(* Logix 5000 project; controller TFF vendor 1 type 14 code 107 rev 34.11; software revision 34.03; part 12 of 36 *)

        LevelConfiguration[0].Alm_HIHITMR := 2, LevelConfiguration[0].Alm_HIHITMR_PRE := 2, LevelConfiguration[1].Alm_HI := 50.0, LevelConfiguration[1].Alm_HI_PRE := 50.0, LevelConfiguration[1].Alm_HIHI := 50.0, LevelConfiguration[1].Alm_HIHI_PRE := 50.0, LevelConfiguration[1].Alm_LOLOTMR := 2, LevelConfiguration[1].Alm_LOLOTMR_PRE := 2, LevelConfiguration[1].Alm_LOTMR := 2, LevelConfiguration[1].Alm_LOTMR_PRE := 2, LevelConfiguration[1].Alm_HITMR := 2, LevelConfiguration[1].Alm_HITMR_PRE := 2, LevelConfiguration[1].Alm_HIHITMR := 2, LevelConfiguration[1].Alm_HIHITMR_PRE := 2, LevelConfiguration[2].Alm_LOLO := 20.0, LevelConfiguration[2].Alm_LOLO_PRE := 20.0, LevelConfiguration[2].Alm_LO := 40.0, LevelConfiguration[2].Alm_LO_PRE := 40.0, LevelConfiguration[2].Alm_HI := 160.0, LevelConfiguration[2].Alm_HI_PRE := 160.0, LevelConfiguration[2].Alm_HIHI := 180.0, LevelConfiguration[2].Alm_HIHI_PRE := 180.0, LevelConfiguration[2].Alm_LOLOTMR := 2, LevelConfiguration[2].Alm_LOLOTMR_PRE := 2, LevelConfiguration[2].Alm_LOTMR := 2, LevelConfiguration[2].Alm_LOTMR_PRE := 2, LevelConfiguration[2].Alm_HITMR := 2, LevelConfiguration[2].Alm_HITMR_PRE := 2, LevelConfiguration[2].Alm_HIHITMR := 2, LevelConfiguration[2].Alm_HIHITMR_PRE := 2, LevelConfiguration[3].Alm_HI := 190.0, LevelConfiguration[3].Alm_HI_PRE := 190.0, LevelConfiguration[3].Alm_HIHI := 200.0, LevelConfiguration[3].Alm_HIHI_PRE := 200.0, Feed_Bag_Tare_Timer.PRE := 3000, Filtrate_Bag_Tare_Timer.PRE := 3000);   // Tank Management
   ThisSystem : SystemType := (Value := 2, MoldType := 124, PreviousValue := 124, EnableSystemType[0] := 1, EnableSystemType[1] := 1, EnableSystemType[2] := 1, EnableSystemType[3] := 1, NewSystem_Timer.PRE := 60000, NewSystem_Timer.ACC := 177455, NewSystem_Timer.EN := 1, NewSystem_Timer.DN := 1);
   TI001 : ALIAS FOR AnalogPoint[13];   // Feed Bag Temperature
   TI001_SIG : ALIAS FOR DigitalPoint[101];
   TI001Alarm : ALIAS FOR AlarmAnalog[13];   // Feed Bag Temperature Alarm
   TimerControl : TimerControl := (Save := 20456, Seconds := 20456, Colon := ':', ColonZero := ':0', Cycle := 818248);   // Timer Control
   Timers : Timers[22] := ([0].TotalSeconds := 30.0, [0].Seconds := 30, [0].sHours := '0', [0].sMinutes := '0', [0].sSeconds := '30', [0].HMS := '0:00:30', [0].LastHMS := '0:02:09', [1].sHours := '0', [1].sMinutes := '0', [1].sSeconds := '0', [1].HMS := '0:00:00', [2].sHours := '0', [2].sMinutes := '0', [2].sSeconds := '0', [2].HMS := '0:00:00', [3].TotalSeconds := 7.0, [3].Seconds := 7, [3].sHours := '0', [3].sMinutes := '0', [3].sSeconds := '7', [3].HMS := '0:00:07', [3].LastHMS := '0:00:00', [4].TotalSeconds := 2.0, [4].Seconds := 2, [4].sHours := '0', [4].sMinutes := '0', [4].sSeconds := '2', [4].HMS := '0:00:02', [5].sHours := '0', [5].sMinutes := '0', [5].sSeconds := '0', [5].HMS := '0:00:00', [5].LastHMS := ':00$00$07$00$00$000:00:00$00$00$00$00$00$00$00$00$00$07$00$00$00', [6].sHours := '0', [6].sMinutes := '0', [6].sSeconds := '0', [6].HMS := '0:00:00', [6].LastHMS := '0:00:02', [7].sHours := '0', [7].sMinutes := '0', [7].sSeconds := '0', [7].HMS := '0:00:00', [8].sHours := '0', [8].sMinutes := '0', [8].sSeconds := '0', [8].HMS := '0:00:00', [8].LastHMS := '$07$00$00$000:00:00$00$00$00$00$00$00$00$00$00$07$00$00$000:$00$00', [9].sHours := '0', [9].sMinutes := '0', [9].sSeconds := '0', [9].HMS := '0:00:00', [9].LastHMS := '$00$00$00$00$00$00$00$00$07$00$00$000:00:00$00$07$00$00$000:$00$00', [10].sHours := '0', [10].sMinutes := '0', [10].sSeconds := '0', [10].HMS := '0:00:00', [10].LastHMS := '0:00:00', [11].sHours := '0', [11].sMinutes := '0', [11].sSeconds := '0',
        [11].HMS := '0:00:00', [11].LastHMS := '0:00:00', [12].sHours := '0', [12].sMinutes := '0', [12].sSeconds := '0', [12].HMS := '0:00:00', [13].TotalSeconds := 16.0, [13].Seconds := 16, [13].sHours := '0', [13].sMinutes := '0', [13].sSeconds := '16', [13].HMS := '0:00:16', [13].LastHMS := ':00$00$07$00$00$000:00:00$00$00$00$00$00$00$00$00$00$07$00$00$00', [14].sHours := '0', [14].sMinutes := '0', [14].sSeconds := '0', [14].HMS := '0:00:00', [14].LastHMS := ':00$00$00$00$00$00$00$00$00$00$07$00$00$000:00:00$00$07$00$00$00', [15].sHours := '0', [15].sMinutes := '0', [15].sSeconds := '0', [15].HMS := '0:00:00', [16].sHours := '0', [16].sMinutes := '0', [16].sSeconds := '0', [16].HMS := '0:00:00', [16].LastHMS := '$07$00$00$000:00:00$00$00$00$00$00$00$00$00$00$07$00$00$000:$00$00', [17].sHours := '0', [17].sMinutes := '0', [17].sSeconds := '0', [17].HMS := '0:00:00', [17].LastHMS := '$00$00$00$00$00$00$00$00$07$00$00$000:00:00$00$07$00$00$000:$00$00', [18].sHours := '0', [18].sMinutes := '0', [18].sSeconds := '0', [18].HMS := '0:00:00', [18].LastHMS := '0:00:00', [19].TotalSeconds := 30.0, [19].Seconds := 30, [19].sHours := '0', [19].sMinutes := '0', [19].sSeconds := '30', [19].HMS := '0:00:30', [19].LastHMS := '0:00:00', [20].sHours := '0', [20].sMinutes := '0', [20].sSeconds := '0', [20].HMS := '0:00:00', [21].sHours := '0', [21].sMinutes := '0', [21].sSeconds := '0', [21].HMS := '0:00:00', [21].LastHMS := '0:00:00');   // Timer Array
        [0]   // Phase 0 Total Time
        [1]   // Phase 1 Total Time
        [2]   // Phase 2 Total Time
        [19]   // Procedure Time
        [3]   // Phase 3 Total Time
        [4]   // Phase 4 Total Time
        [10]   // Phase 4 Step Time
        [11]   // Phase 5 Step Time
        [5]   // Phase 5 Total Time
        [12]   // Phase 0 Pause Time
        [13]   // Phase 1 Pause Time
        [14]   // Phase 2 Pause Time
        [15]   // Phase 3 Pause Time
        [16]   // Phase 4 Pause Time
        [17]   // Phase 5 Pause Time
        [18]   // User Time
        [21]   // Linear Gradient
        [6]   // Phase 0 Step Time
        [7]   // Phase 1 Step Time
        [8]   // Phase 2 Step Time
        [9]   // Phase 3 Step Time
   TMP : ALIAS FOR AnalogPoint[41];   // Trans-membrane Pressure
   TMPAlarm : ALIAS FOR AlarmAnalog[41];   // Trans-membrane Pressure Alarm
   Totalizer : Totalizers[20] := ([0].PVscale := 60.0, [0].Title := 'Conc', [0].ResetTimer.PRE := 3000, [1].PVscale := 60.0, [1].Title := 'Diaf', [1].ResetTimer.PRE := 3000, [2].PVsec := inf, [2].ResetTimer.PRE := 3000, [3].PVsec := inf, [3].ResetTimer.PRE := 3000, [4].ResetTimer.PRE := 3000, [5].ResetTimer.PRE := 3000, [6].ResetTimer.PRE := 3000, [7].ResetTimer.PRE := 3000, [8].ResetTimer.PRE := 3000, [9].ResetTimer.PRE := 3000, [10].ResetTimer.PRE := 3000, [11].ResetTimer.PRE := 3000, [12].ResetTimer.PRE := 3000, [13].ResetTimer.PRE := 3000, [14].ResetTimer.PRE := 3000, [15].ResetTimer.PRE := 3000, [16].ResetTimer.PRE := 3000, [17].ResetTimer.PRE := 3000, [18].ResetTimer.PRE := 3000, [19].ResetTimer.PRE := 3000);   // Totalizers Array
        [0]   // Concentration totalizer
        [1]   // Diafiltration totalizer
   Transfer_Pump_P002_Type : INT := 1;   // Transfer Pump P002 Type Status
   UserAlarm : UserAlarm;   // User Alarm (used in CCP Recipe)
   UserCr1 : ALIAS FOR DigitalPoint[65];   // User Critical Alarm 1
   UserCr2 : ALIAS FOR DigitalPoint[67];   // User Critical Alarm 2
   UserNCr1 : ALIAS FOR DigitalPoint[64];   // User Non Critical Alarm 1
   UserNCr2 : ALIAS FOR DigitalPoint[66];   // User Non Critical Alarm 2
   UserTime : ALIAS FOR Timers[18];   // User time
   UserTotalizerManagement : UserTotalizerManagement := (LogUserTimer.PRE := 3000, ResetUserTimer.PRE := 3000);   // User Totalizer management
   Valve : Valve[100] := ([0].Tag := 'XV001', [0].Control := 1, [0].Auto := 1, [0].Manual := 1, [0].OpenStatus := 1, [0].ZSOverride := 1, [0].FailState := 1, [0].EnableCfg := 1, [0].StatusWord := 2, [0].Status := 2, [0].OutputAddress := 32, [0].AlarmTimer.PRE := 2000, [0].AlarmTimerSP := 2, [1].Tag := 'XV002', [1].Control := 1, [1].Auto := 1, [1].Manual := 1, [1].OpenStatus := 1, [1].ZSOverride := 1, [1].FailState := 1, [1].EnableCfg := 1, [1].StatusWord := 2, [1].Status := 2, [1].OutputAddress := 33, [1].AlarmTimer.PRE := 2000, [1].AlarmTimerSP := 2, [1].AutoCloseTimer.ACC := 1103, [2].Tag := 'XV003', [2].Control := 1, [2].Auto := 1, [2].Manual := 1, [2].OpenStatus := 1, [2].ZSOverride := 1, [2].EnableCfg := 1, [2].StatusWord := 2, [2].Status := 2, [2].OutputAddress := 34, [2].AlarmTimer.PRE := 2000, [2].AlarmTimerSP := 2, [2].AutoCloseTimer.ACC := 1032, [3].Tag := 'XV004', [3].Control := 1, [3].Auto := 1, [3].Manual := 1, [3].OpenStatus := 1, [3].ZSOverride := 1, [3].FailState := 1, [3].EnableCfg := 1, [3].StatusWord := 2, [3].Status := 2, [3].OutputAddress := 35, [3].AlarmTimer.PRE := 2000, [3].AlarmTimerSP := 2, [3].AutoCloseTimer.ACC := 1115, [4].Tag := 'XV005', [4].Control := 1, [4].Auto := 1, [4].Manual := 1, [4].OpenStatus := 1, [4].ZSOverride := 1,
        [4].EnableCfg := 1, [4].StatusWord := 2, [4].Status := 2, [4].OutputAddress := 36, [4].AlarmTimer.PRE := 2000, [4].AlarmTimerSP := 2, [4].AutoCloseTimer.ACC := 1104, [5].Tag := 'XV102', [5].Control := 1, [5].Auto := 1, [5].Manual := 1, [5].OpenStatus := 1, [5].ZSOverride := 1, [5].EnableCfg := 1, [5].StatusWord := 2, [5].Status := 2, [5].OutputAddress := 38, [5].AlarmTimer.PRE := 2000, [5].AlarmTimerSP := 2, [5].AutoCloseTimer.ACC := 1104, [6].Tag := 'XV401', [6].Control := 1, [6].Auto := 1, [6].Manual := 1, [6].OpenStatus := 1, [6].ZSOverride := 1, [6].EnableCfg := 1, [6].StatusWord := 2, [6].Status := 2, [6].OutputAddress := 41, [6].AlarmTimer.PRE := 2000, [6].AlarmTimerSP := 2, [6].AutoCloseTimer.ACC := 1104, [7].Tag := 'XV402', [7].CloseStatus := 1, [7].ZSOverride := 1, [7].EnableCfg := 1, [7].StatusWord := 4, [7].Status := 4, [7].OutputAddress := 42, [7].AlarmTimer.PRE := 2000, [7].AlarmTimerSP := 2, [7].AutoCloseTimer.ACC := 1104, [8].Tag := 'XV411', [8].CloseStatus := 1, [8].ZSOverride := 1, [8].EnableCfg := 1, [8].StatusWord := 4, [8].Status := 4, [8].OutputAddress := 43, [8].AlarmTimer.PRE := 2000, [8].AlarmTimerSP := 2, [8].AutoCloseTimer.ACC := 1104, [9].Tag := 'XV421', [9].CloseStatus := 1, [9].ZSOverride := 1, [9].EnableCfg := 1, [9].StatusWord := 4, [9].Status := 4, [9].OutputAddress := 44,
        [9].AlarmTimer.PRE := 2000, [9].AlarmTimerSP := 2, [9].AutoCloseTimer.ACC := 1105, [10].Tag := 'XV431', [10].CloseStatus := 1, [10].ZSOverride := 1, [10].EnableCfg := 1, [10].StatusWord := 4, [10].Status := 4, [10].OutputAddress := 45, [10].AlarmTimer.PRE := 2000, [10].AlarmTimerSP := 2, [10].AutoCloseTimer.ACC := 1104, [11].Tag := 'XV441', [11].Control := 1, [11].Auto := 1, [11].Manual := 1, [11].OpenStatus := 1, [11].ZSOverride := 1, [11].EnableCfg := 1, [11].StatusWord := 2, [11].Status := 2, [11].OutputAddress := 46, [11].AlarmTimer.PRE := 2000, [11].AlarmTimerSP := 2, [11].AutoCloseTimer.ACC := 1103, [12].Tag := 'XV501', [12].Control := 1, [12].Auto := 1, [12].Manual := 1, [12].OpenStatus := 1, [12].ZSOverride := 1, [12].EnableCfg := 1, [12].StatusWord := 2, [12].Status := 2, [12].OutputAddress := 39, [12].AlarmTimer.PRE := 2000, [12].AlarmTimerSP := 2, [12].AutoCloseTimer.ACC := 1072, [13].Tag := 'XV502', [13].Control := 1, [13].Auto := 1, [13].Manual := 1, [13].OpenStatus := 1, [13].ZSOverride := 1, [13].EnableCfg := 1, [13].StatusWord := 2, [13].Status := 2, [13].OutputAddress := 40, [13].AlarmTimer.PRE := 2000, [13].AlarmTimerSP := 2, [13].AutoCloseTimer.ACC := 1016, [14].Tag := 'XV901', [14].Control := 1, [14].Auto := 1, [14].Manual := 1, [14].OpenStatus := 1, [14].ZSOverride := 1, [14].EnableCfg := 1, [14].StatusWord := 2,
        [14].Status := 2, [14].OutputAddress := 37, [14].AlarmTimer.PRE := 2000, [14].AlarmTimerSP := 2, [15].OpenStatus := 1, [15].ZSOverride := 1, [15].OutputAddress := 47, [15].AlarmTimer.PRE := 2000, [15].AlarmTimerSP := 2, [16].CloseStatus := 1, [16].ZSOverride := 1, [16].OutputAddress := 48, [16].AlarmTimer.PRE := 2000, [16].AlarmTimerSP := 2, [17].OpenStatus := 1, [17].ZSOverride := 1, [17].OutputAddress := 49, [17].AlarmTimer.PRE := 2000, [17].AlarmTimerSP := 2, [17].AutoCloseTimer.ACC := 1594, [18].CloseStatus := 1, [18].ZSOverride := 1, [18].OutputAddress := 50, [18].AlarmTimer.PRE := 2000, [18].AlarmTimerSP := 2, [18].AutoCloseTimer.ACC := 137, [19].CloseStatus := 1, [19].ZSOverride := 1, [19].FailState := 1, [19].OutputAddress := 51, [19].AlarmTimer.PRE := 2000, [19].AlarmTimerSP := 2, [19].AutoCloseTimer.ACC := 1007, [20].CloseStatus := 1, [20].ZSOverride := 1, [20].OutputAddress := 52, [20].AlarmTimer.PRE := 2000, [20].AlarmTimerSP := 2, [20].AutoCloseTimer.ACC := 1004, [21].OpenStatus := 1, [21].ZSOverride := 1, [21].FailState := 1, [21].OutputAddress := 53, [21].AlarmTimer.PRE := 2000, [21].AlarmTimerSP := 2, [22].CloseStatus := 1, [22].ZSOverride := 1, [22].OutputAddress := 54, [22].AlarmTimer.PRE := 2000, [22].AlarmTimerSP := 2, [22].AutoCloseTimer.ACC := 131, [23].CloseStatus := 1, [23].ZSOverride := 1, [23].OutputAddress := 55, [23].AlarmTimer.PRE := 2000, [23].AlarmTimerSP := 2, [23].AutoCloseTimer.ACC := 1003, [24].CloseStatus := 1, [24].ZSOverride := 1, [24].OutputAddress := 56,
        [24].AlarmTimer.PRE := 2000, [24].AlarmTimerSP := 2, [24].AutoCloseTimer.ACC := 1002, [25].CloseStatus := 1, [25].ZSOverride := 1, [25].OutputAddress := 57, [25].AlarmTimer.PRE := 2000, [25].AlarmTimerSP := 2, [25].AutoCloseTimer.ACC := 1002, [26].CloseStatus := 1, [26].ZSOverride := 1, [26].OutputAddress := 58, [26].AlarmTimer.PRE := 2000, [26].AlarmTimerSP := 2, [26].AutoCloseTimer.ACC := 1002, [27].CloseStatus := 1, [27].ZSOverride := 1, [27].OutputAddress := 59, [27].AlarmTimer.PRE := 2000, [27].AlarmTimerSP := 2, [28].CloseStatus := 1, [28].ZSOverride := 1, [28].OutputAddress := 60, [28].AlarmTimer.PRE := 2000, [28].AlarmTimerSP := 2, [29].OpenStatus := 1, [29].ZSOverride := 1, [29].FailState := 1, [29].OutputAddress := 61, [29].AlarmTimer.PRE := 2000, [29].AlarmTimerSP := 2, [29].AutoCloseTimer.ACC := 1068, [30].CloseStatus := 1, [30].ZSOverride := 1, [30].OutputAddress := 62, [30].AlarmTimer.PRE := 2000, [30].AlarmTimerSP := 2, [30].AutoCloseTimer.ACC := 1069, [31].CloseStatus := 1, [31].ZSOverride := 1, [31].OutputAddress := 63, [31].AlarmTimer.PRE := 2000, [31].AlarmTimerSP := 2, [31].AutoCloseTimer.ACC := 131, [32].CloseStatus := 1, [32].PriorityCfg := 1, [32].AlarmTimerSP := 2, [32].AutoCloseTimer.ACC := 1059, [33].OpenStatus := 1, [33].PriorityCfg := 1, [33].AlarmTimerSP := 2, [33].AutoCloseTimer.ACC := 1123, [34].OpenStatus := 1, [34].PriorityCfg := 1, [34].AlarmTimerSP := 2, [34].AutoCloseTimer.ACC := 1095, [35].OpenStatus := 1, [35].PriorityCfg := 1, [35].AlarmTimerSP := 2, [35].AutoCloseTimer.ACC := 1127,
        [36].OpenStatus := 1, [36].PriorityCfg := 1, [36].AlarmTimerSP := 2, [36].AutoCloseTimer.ACC := 1004, [37].CloseStatus := 1, [37].PriorityCfg := 1, [37].AlarmTimerSP := 2, [37].AutoCloseTimer.ACC := 1121, [38].CloseStatus := 1, [38].Priority := 1, [38].PriorityCfg := 1, [38].AlarmTimerSP := 2, [38].AutoCloseTimer.ACC := 1135, [39].CloseStatus := 1, [39].Priority := 1, [39].PriorityCfg := 1, [39].AlarmTimerSP := 2, [39].AutoCloseTimer.ACC := 1121, [40].CloseStatus := 1, [40].Priority := 1, [40].PriorityCfg := 1, [40].AlarmTimerSP := 2, [40].AutoCloseTimer.ACC := 1112, [41].CloseStatus := 1, [41].Priority := 1, [41].PriorityCfg := 1, [41].AlarmTimerSP := 2, [42].CloseStatus := 1, [42].Priority := 1, [42].PriorityCfg := 1, [42].AlarmTimerSP := 2, [43].CloseStatus := 1, [43].Priority := 1, [43].PriorityCfg := 1, [43].AlarmTimerSP := 2, [44].CloseStatus := 1, [44].Priority := 1, [44].PriorityCfg := 1, [44].AlarmTimerSP := 2, [45].CloseStatus := 1, [45].Priority := 1, [45].PriorityCfg := 1, [45].AlarmTimerSP := 2, [46].CloseStatus := 1, [46].Priority := 1, [46].PriorityCfg := 1, [46].AlarmTimerSP := 2, [47].OpenStatus := 1, [47].Priority := 1, [47].PriorityCfg := 1, [47].AlarmTimerSP := 2, [51].OpenStatus := 1, [52].OpenStatus := 1, [53].CloseStatus := 1, [54].CloseStatus := 1, [55].CloseStatus := 1, [56].CloseStatus := 1, [58].CloseStatus := 1, [59].CloseStatus := 1);   // Valve Array
        [10]   // XV431
        [11]   // XV441
        [12]   // XV501
        [13]   // XV502
        [14]   // XV901
        [15]   // XV403
        [16]   // XV404
        [17]   // XV405
        [18]   // XV406
        [0]   // XV001
        [19]   // XV006
        [1]   // XV002
        [20]   // XV007
        [2]   // XV003
        [0].FailState   // Valve Fail State 0=Closed 1=Open
        [3]   // XV004
        [4]   // XV005
        [5]   // XV102
        [6]   // XV401
        [7]   // XV402
        [8]   // XV411
        [9]   // XV421
   Valve_Storage : Valve[6,100] := ([0,0].Tag := 'XV001', [0,0].CloseStatus := 1, [0,0].ZSOverride := 1, [0,0].EnableCfg := 1, [0,0].StatusWord := 4, [0,0].Status := 4, [0,0].OutputAddress := 32, [0,0].AlarmTimer.PRE := 2000, [0,0].AlarmTimerSP := 2, [0,1].Tag := 'XV002', [0,1].CloseStatus := 1, [0,1].ZSOverride := 1, [0,1].EnableCfg := 1, [0,1].StatusWord := 4, [0,1].Status := 4, [0,1].OutputAddress := 33, [0,1].AlarmTimer.PRE := 2000, [0,1].AlarmTimerSP := 2, [0,1].AutoCloseTimer.ACC := 1103, [0,2].Tag := 'XV003', [0,2].CloseStatus := 1, [0,2].ZSOverride := 1, [0,2].EnableCfg := 1, [0,2].StatusWord := 4, [0,2].Status := 4, [0,2].OutputAddress := 34, [0,2].AlarmTimer.PRE := 2000, [0,2].AlarmTimerSP := 2, [0,2].AutoCloseTimer.ACC := 1032, [0,3].Tag := 'XV004', [0,3].CloseStatus := 1, [0,3].ZSOverride := 1, [0,3].EnableCfg := 1, [0,3].StatusWord := 4, [0,3].Status := 4, [0,3].OutputAddress := 35, [0,3].AlarmTimer.PRE := 2000, [0,3].AlarmTimerSP := 2, [0,3].AutoCloseTimer.ACC := 1115, [0,4].Tag := 'XV005', [0,4].CloseStatus := 1, [0,4].ZSOverride := 1, [0,4].EnableCfg := 1, [0,4].StatusWord := 4, [0,4].Status := 4, [0,4].OutputAddress := 36, [0,4].AlarmTimer.PRE := 2000, [0,4].AlarmTimerSP := 2, [0,4].AutoCloseTimer.ACC := 1104, [0,5].Tag := 'XV006', [0,5].CloseStatus := 1, [0,5].ZSOverride := 1, [0,5].EnableCfg := 1, [0,5].StatusWord := 4, [0,5].Status := 4, [0,5].OutputAddress := 37, [0,5].AlarmTimer.PRE := 2000, [0,5].AlarmTimerSP := 2, [0,5].AutoCloseTimer.ACC := 1104, [0,6].Tag := 'XV007',
        [0,6].CloseStatus := 1, [0,6].ZSOverride := 1, [0,6].EnableCfg := 1, [0,6].StatusWord := 4, [0,6].Status := 4, [0,6].OutputAddress := 38, [0,6].AlarmTimer.PRE := 2000, [0,6].AlarmTimerSP := 2, [0,6].AutoCloseTimer.ACC := 1104, [0,7].Tag := 'XV008', [0,7].CloseStatus := 1, [0,7].ZSOverride := 1, [0,7].EnableCfg := 1, [0,7].StatusWord := 4, [0,7].Status := 4, [0,7].OutputAddress := 39, [0,7].AlarmTimer.PRE := 2000, [0,7].AlarmTimerSP := 2, [0,7].AutoCloseTimer.ACC := 1104, [0,8].Tag := 'XV009', [0,8].CloseStatus := 1, [0,8].ZSOverride := 1, [0,8].EnableCfg := 1, [0,8].StatusWord := 4, [0,8].Status := 4, [0,8].OutputAddress := 40, [0,8].AlarmTimer.PRE := 2000, [0,8].AlarmTimerSP := 2, [0,8].AutoCloseTimer.ACC := 1104, [0,9].Tag := 'XV010', [0,9].CloseStatus := 1, [0,9].ZSOverride := 1, [0,9].EnableCfg := 1, [0,9].StatusWord := 4, [0,9].Status := 4, [0,9].OutputAddress := 41, [0,9].AlarmTimer.PRE := 2000, [0,9].AlarmTimerSP := 2, [0,9].AutoCloseTimer.ACC := 1105, [0,10].Tag := 'XV011', [0,10].CloseStatus := 1, [0,10].ZSOverride := 1, [0,10].EnableCfg := 1, [0,10].StatusWord := 4, [0,10].Status := 4, [0,10].OutputAddress := 42, [0,10].AlarmTimer.PRE := 2000, [0,10].AlarmTimerSP := 2, [0,10].AutoCloseTimer.ACC := 1104, [0,11].Tag := 'XV012', [0,11].Control := 1, [0,11].Auto := 1, [0,11].Manual := 1, [0,11].OpenStatus := 1, [0,11].ZSOverride := 1, [0,11].FailState := 1, [0,11].EnableCfg := 1, [0,11].StatusWord := 2, [0,11].Status := 2, [0,11].OutputAddress := 43,
        [0,11].AlarmTimer.PRE := 2000, [0,11].AlarmTimerSP := 2, [0,11].AutoCloseTimer.ACC := 1103, [0,12].Tag := 'XV013', [0,12].Control := 1, [0,12].Auto := 1, [0,12].Manual := 1, [0,12].OpenStatus := 1, [0,12].ZSOverride := 1, [0,12].FailState := 1, [0,12].EnableCfg := 1, [0,12].StatusWord := 2, [0,12].Status := 2, [0,12].OutputAddress := 44, [0,12].AlarmTimer.PRE := 2000, [0,12].AlarmTimerSP := 2, [0,12].AutoCloseTimer.ACC := 1072, [0,13].Tag := 'XV014', [0,13].Control := 1, [0,13].Auto := 1, [0,13].Manual := 1, [0,13].OpenStatus := 1, [0,13].ZSOverride := 1, [0,13].FailState := 1, [0,13].EnableCfg := 1, [0,13].StatusWord := 2, [0,13].Status := 2, [0,13].OutputAddress := 45, [0,13].AlarmTimer.PRE := 2000, [0,13].AlarmTimerSP := 2, [0,13].AutoCloseTimer.ACC := 1016, [0,14].Tag := 'XV015', [0,14].CloseStatus := 1, [0,14].ZSOverride := 1, [0,14].EnableCfg := 1, [0,14].StatusWord := 4, [0,14].Status := 4, [0,14].OutputAddress := 46, [0,14].AlarmTimer.PRE := 2000, [0,14].AlarmTimerSP := 2, [0,15].Tag := 'XV016', [0,15].Control := 1, [0,15].Auto := 1, [0,15].Manual := 1, [0,15].OpenStatus := 1, [0,15].ZSOverride := 1, [0,15].FailState := 1, [0,15].EnableCfg := 1, [0,15].StatusWord := 2, [0,15].Status := 2, [0,15].OutputAddress := 47, [0,15].AlarmTimer.PRE := 2000, [0,15].AlarmTimerSP := 2, [0,16].Tag := 'XV017', [0,16].CloseStatus := 1, [0,16].ZSOverride := 1, [0,16].EnableCfg := 1, [0,16].StatusWord := 4, [0,16].Status := 4, [0,16].OutputAddress := 48,
        [0,16].AlarmTimer.PRE := 2000, [0,16].AlarmTimerSP := 2, [0,17].Tag := 'XV018', [0,17].Control := 1, [0,17].Auto := 1, [0,17].Manual := 1, [0,17].OpenStatus := 1, [0,17].ZSOverride := 1, [0,17].FailState := 1, [0,17].EnableCfg := 1, [0,17].StatusWord := 2, [0,17].Status := 2, [0,17].OutputAddress := 49, [0,17].AlarmTimer.PRE := 2000, [0,17].AlarmTimerSP := 2, [0,17].AutoCloseTimer.ACC := 1594, [0,18].Tag := 'XV019', [0,18].CloseStatus := 1, [0,18].ZSOverride := 1, [0,18].EnableCfg := 1, [0,18].StatusWord := 4, [0,18].Status := 4, [0,18].OutputAddress := 50, [0,18].AlarmTimer.PRE := 2000, [0,18].AlarmTimerSP := 2, [0,18].AutoCloseTimer.ACC := 137, [0,19].Tag := 'XV020', [0,19].CloseStatus := 1, [0,19].ZSOverride := 1, [0,19].EnableCfg := 1, [0,19].StatusWord := 4, [0,19].Status := 4, [0,19].OutputAddress := 51, [0,19].AlarmTimer.PRE := 2000, [0,19].AlarmTimerSP := 2, [0,19].AutoCloseTimer.ACC := 1007, [0,20].Tag := 'XV021', [0,20].CloseStatus := 1, [0,20].ZSOverride := 1, [0,20].EnableCfg := 1, [0,20].StatusWord := 4, [0,20].Status := 4, [0,20].OutputAddress := 52, [0,20].AlarmTimer.PRE := 2000, [0,20].AlarmTimerSP := 2, [0,20].AutoCloseTimer.ACC := 1004, [0,21].Tag := 'XV022', [0,21].Control := 1, [0,21].Auto := 1, [0,21].Manual := 1, [0,21].OpenStatus := 1, [0,21].ZSOverride := 1, [0,21].FailState := 1, [0,21].EnableCfg := 1, [0,21].StatusWord := 2, [0,21].Status := 2, [0,21].OutputAddress := 53, [0,21].AlarmTimer.PRE := 2000, [0,21].AlarmTimerSP := 2, [0,22].Tag := 'XV023',
        [0,22].CloseStatus := 1, [0,22].ZSOverride := 1, [0,22].EnableCfg := 1, [0,22].StatusWord := 4, [0,22].Status := 4, [0,22].OutputAddress := 54, [0,22].AlarmTimer.PRE := 2000, [0,22].AlarmTimerSP := 2, [0,22].AutoCloseTimer.ACC := 131, [0,23].Tag := 'XV024', [0,23].CloseStatus := 1, [0,23].ZSOverride := 1, [0,23].EnableCfg := 1, [0,23].StatusWord := 4, [0,23].Status := 4, [0,23].OutputAddress := 55, [0,23].AlarmTimer.PRE := 2000, [0,23].AlarmTimerSP := 2, [0,23].AutoCloseTimer.ACC := 1003, [0,24].Tag := 'XV025', [0,24].CloseStatus := 1, [0,24].ZSOverride := 1, [0,24].EnableCfg := 1, [0,24].StatusWord := 4, [0,24].Status := 4, [0,24].OutputAddress := 56, [0,24].AlarmTimer.PRE := 2000, [0,24].AlarmTimerSP := 2, [0,24].AutoCloseTimer.ACC := 1002, [0,25].Tag := 'XV026', [0,25].CloseStatus := 1, [0,25].ZSOverride := 1, [0,25].EnableCfg := 1, [0,25].StatusWord := 4, [0,25].Status := 4, [0,25].OutputAddress := 57, [0,25].AlarmTimer.PRE := 2000, [0,25].AlarmTimerSP := 2, [0,25].AutoCloseTimer.ACC := 1002, [0,26].Tag := 'XV028', [0,26].CloseStatus := 1, [0,26].ZSOverride := 1, [0,26].EnableCfg := 1, [0,26].StatusWord := 4, [0,26].Status := 4, [0,26].OutputAddress := 58, [0,26].AlarmTimer.PRE := 2000, [0,26].AlarmTimerSP := 2, [0,26].AutoCloseTimer.ACC := 1002, [0,27].Tag := 'XV029', [0,27].CloseStatus := 1, [0,27].ZSOverride := 1, [0,27].EnableCfg := 1, [0,27].StatusWord := 4, [0,27].Status := 4, [0,27].OutputAddress := 59, [0,27].AlarmTimer.PRE := 2000, [0,27].AlarmTimerSP := 2, [0,28].Tag := 'XV030', [0,28].CloseStatus := 1,
        [0,28].ZSOverride := 1, [0,28].EnableCfg := 1, [0,28].StatusWord := 4, [0,28].Status := 4, [0,28].OutputAddress := 60, [0,28].AlarmTimer.PRE := 2000, [0,28].AlarmTimerSP := 2, [0,29].Tag := 'XV031', [0,29].Control := 1, [0,29].Auto := 1, [0,29].Manual := 1, [0,29].OpenStatus := 1, [0,29].ZSOverride := 1, [0,29].FailState := 1, [0,29].EnableCfg := 1, [0,29].StatusWord := 2, [0,29].Status := 2, [0,29].OutputAddress := 61, [0,29].AlarmTimer.PRE := 2000, [0,29].AlarmTimerSP := 2, [0,29].AutoCloseTimer.ACC := 1068, [0,30].Tag := 'XV033', [0,30].CloseStatus := 1, [0,30].ZSOverride := 1, [0,30].EnableCfg := 1, [0,30].StatusWord := 4, [0,30].Status := 4, [0,30].OutputAddress := 62, [0,30].AlarmTimer.PRE := 2000, [0,30].AlarmTimerSP := 2, [0,30].AutoCloseTimer.ACC := 1069, [0,31].Tag := 'XV034', [0,31].CloseStatus := 1, [0,31].ZSOverride := 1, [0,31].EnableCfg := 1, [0,31].StatusWord := 4, [0,31].Status := 4, [0,31].OutputAddress := 63, [0,31].AlarmTimer.PRE := 2000, [0,31].AlarmTimerSP := 2, [0,31].AutoCloseTimer.ACC := 131, [0,32].CloseStatus := 1, [0,32].PriorityCfg := 1, [0,32].ZSOpenAddress := 32, [0,32].OutputAddress := 68, [0,32].AlarmTimer.PRE := 2000, [0,32].AlarmTimerSP := 2, [0,32].AutoCloseTimer.ACC := 1059, [0,33].OpenStatus := 1, [0,33].PriorityCfg := 1, [0,33].FailState := 1, [0,33].ZSCloseAddress := 33, [0,33].OutputAddress := 69, [0,33].AlarmTimer.PRE := 2000, [0,33].AlarmTimerSP := 2, [0,33].AutoCloseTimer.ACC := 1123, [0,34].OpenStatus := 1, [0,34].PriorityCfg := 1, [0,34].FailState := 1, [0,34].ZSCloseAddress := 34,
        [0,34].OutputAddress := 70, [0,34].AlarmTimer.PRE := 2000, [0,34].AlarmTimerSP := 2, [0,34].AutoCloseTimer.ACC := 1095, [0,35].OpenStatus := 1, [0,35].PriorityCfg := 1, [0,35].FailState := 1, [0,35].ZSCloseAddress := 35, [0,35].OutputAddress := 71, [0,35].AlarmTimer.PRE := 2000, [0,35].AlarmTimerSP := 2, [0,35].AutoCloseTimer.ACC := 1127, [0,36].OpenStatus := 1, [0,36].PriorityCfg := 1, [0,36].FailState := 1, [0,36].ZSCloseAddress := 36, [0,36].OutputAddress := 72, [0,36].AlarmTimer.PRE := 2000, [0,36].AlarmTimerSP := 2, [0,36].AutoCloseTimer.ACC := 1004, [0,37].CloseStatus := 1, [0,37].PriorityCfg := 1, [0,37].ZSOpenAddress := 37, [0,37].OutputAddress := 73, [0,37].AlarmTimer.PRE := 2000, [0,37].AlarmTimerSP := 2, [0,37].AutoCloseTimer.ACC := 1121, [0,38].CloseStatus := 1, [0,38].Priority := 1, [0,38].PriorityCfg := 1, [0,38].ZSOpenAddress := 38, [0,38].OutputAddress := 40, [0,38].AlarmTimer.PRE := 2000, [0,38].AlarmTimerSP := 2, [0,38].AutoCloseTimer.ACC := 1135, [0,39].CloseStatus := 1, [0,39].Priority := 1, [0,39].PriorityCfg := 1, [0,39].ZSOpenAddress := 39, [0,39].OutputAddress := 41, [0,39].AlarmTimer.PRE := 2000, [0,39].AlarmTimerSP := 2, [0,39].AutoCloseTimer.ACC := 1121, [0,40].CloseStatus := 1, [0,40].Priority := 1, [0,40].PriorityCfg := 1, [0,40].ZSOpenAddress := 40, [0,40].OutputAddress := 42, [0,40].AlarmTimer.PRE := 2000, [0,40].AlarmTimerSP := 2, [0,40].AutoCloseTimer.ACC := 1112, [0,41].CloseStatus := 1, [0,41].Priority := 1, [0,41].PriorityCfg := 1, [0,41].ZSOpenAddress := 41, [0,41].OutputAddress := 43, [0,41].AlarmTimer.PRE := 2000, [0,41].AlarmTimerSP := 2, [0,42].CloseStatus := 1, [0,42].Priority := 1,
        [0,42].PriorityCfg := 1, [0,42].ZSOpenAddress := 42, [0,42].OutputAddress := 44, [0,42].AlarmTimer.PRE := 2000, [0,42].AlarmTimerSP := 2, [0,43].CloseStatus := 1, [0,43].Priority := 1, [0,43].PriorityCfg := 1, [0,43].ZSOpenAddress := 43, [0,43].OutputAddress := 52, [0,43].AlarmTimer.PRE := 2000, [0,43].AlarmTimerSP := 2, [0,44].CloseStatus := 1, [0,44].Priority := 1, [0,44].PriorityCfg := 1, [0,44].ZSOpenAddress := 44, [0,44].OutputAddress := 53, [0,44].AlarmTimer.PRE := 2000, [0,44].AlarmTimerSP := 2, [0,45].CloseStatus := 1, [0,45].Priority := 1, [0,45].PriorityCfg := 1, [0,45].ZSOpenAddress := 45, [0,45].OutputAddress := 54, [0,45].AlarmTimer.PRE := 2000, [0,45].AlarmTimerSP := 2, [0,46].CloseStatus := 1, [0,46].Priority := 1, [0,46].PriorityCfg := 1, [0,46].ZSOpenAddress := 46, [0,46].OutputAddress := 55, [0,46].AlarmTimer.PRE := 2000, [0,46].AlarmTimerSP := 2, [0,47].OpenStatus := 1, [0,47].Priority := 1, [0,47].PriorityCfg := 1, [0,47].FailState := 1, [0,47].ZSCloseAddress := 47, [0,47].OutputAddress := 45, [0,47].AlarmTimer.PRE := 2000, [0,47].AlarmTimerSP := 2, [0,48].FailState := 1, [0,48].ZSCloseAddress := 48, [0,48].OutputAddress := 80, [0,49].FailState := 1, [0,49].ZSCloseAddress := 49, [0,49].OutputAddress := 81, [0,50].FailState := 1, [0,50].ZSCloseAddress := 50, [0,50].OutputAddress := 82, [0,51].OpenStatus := 1, [0,51].FailState := 1, [0,51].ZSCloseAddress := 51, [0,51].OutputAddress := 83, [0,52].OpenStatus := 1, [0,52].FailState := 1, [0,52].ZSCloseAddress := 52, [0,52].OutputAddress := 84, [0,53].CloseStatus := 1, [0,53].FailState := 1,
        [0,53].ZSCloseAddress := 53, [0,53].OutputAddress := 85, [0,54].CloseStatus := 1, [0,54].FailState := 1, [0,54].ZSCloseAddress := 54, [0,54].OutputAddress := 86, [0,55].CloseStatus := 1, [0,55].FailState := 1, [0,55].ZSCloseAddress := 55, [0,55].OutputAddress := 87, [0,56].CloseStatus := 1, [0,58].CloseStatus := 1, [0,59].CloseStatus := 1, [1,0].Tag := 'XV001', [1,0].Control := 1, [1,0].Auto := 1, [1,0].Manual := 1, [1,0].OpenStatus := 1, [1,0].ZSOverride := 1, [1,0].FailState := 1, [1,0].EnableCfg := 1, [1,0].StatusWord := 2, [1,0].Status := 2, [1,0].OutputAddress := 32, [1,0].AlarmTimer.PRE := 2000, [1,0].AlarmTimerSP := 2, [1,1].Tag := 'XV002', [1,1].Control := 1, [1,1].Auto := 1, [1,1].Manual := 1, [1,1].OpenStatus := 1, [1,1].ZSOverride := 1, [1,1].FailState := 1, [1,1].EnableCfg := 1, [1,1].StatusWord := 2, [1,1].Status := 2, [1,1].OutputAddress := 33, [1,1].AlarmTimer.PRE := 2000, [1,1].AlarmTimerSP := 2, [1,1].AutoCloseTimer.ACC := 1103, [1,2].Tag := 'XV003', [1,2].CloseStatus := 1, [1,2].ZSOverride := 1, [1,2].EnableCfg := 1, [1,2].StatusWord := 4, [1,2].Status := 4, [1,2].OutputAddress := 34, [1,2].AlarmTimer.PRE := 2000, [1,2].AlarmTimerSP := 2, [1,2].AutoCloseTimer.ACC := 1032, [1,3].Tag := 'XV004', [1,3].Control := 1, [1,3].Auto := 1, [1,3].Manual := 1, [1,3].OpenStatus := 1, [1,3].ZSOverride := 1, [1,3].FailState := 1, [1,3].EnableCfg := 1, [1,3].StatusWord := 2, [1,3].Status := 2,
        [1,3].OutputAddress := 35, [1,3].AlarmTimer.PRE := 2000, [1,3].AlarmTimerSP := 2, [1,3].AutoCloseTimer.ACC := 1115, [1,4].Tag := 'XV005', [1,4].CloseStatus := 1, [1,4].ZSOverride := 1, [1,4].EnableCfg := 1, [1,4].StatusWord := 4, [1,4].Status := 4, [1,4].OutputAddress := 36, [1,4].AlarmTimer.PRE := 2000, [1,4].AlarmTimerSP := 2, [1,4].AutoCloseTimer.ACC := 1104, [1,5].Tag := 'XV102', [1,5].CloseStatus := 1, [1,5].ZSOverride := 1, [1,5].EnableCfg := 1, [1,5].StatusWord := 4, [1,5].Status := 4, [1,5].OutputAddress := 38, [1,5].AlarmTimer.PRE := 2000, [1,5].AlarmTimerSP := 2, [1,5].AutoCloseTimer.ACC := 1104, [1,6].Tag := 'XV401', [1,6].CloseStatus := 1, [1,6].ZSOverride := 1, [1,6].EnableCfg := 1, [1,6].StatusWord := 4, [1,6].Status := 4, [1,6].OutputAddress := 41, [1,6].AlarmTimer.PRE := 2000, [1,6].AlarmTimerSP := 2, [1,6].AutoCloseTimer.ACC := 1104, [1,7].Tag := 'XV402', [1,7].CloseStatus := 1, [1,7].ZSOverride := 1, [1,7].EnableCfg := 1, [1,7].StatusWord := 4, [1,7].Status := 4, [1,7].OutputAddress := 42, [1,7].AlarmTimer.PRE := 2000, [1,7].AlarmTimerSP := 2, [1,7].AutoCloseTimer.ACC := 1104, [1,8].Tag := 'XV411', [1,8].CloseStatus := 1, [1,8].ZSOverride := 1, [1,8].EnableCfg := 1, [1,8].StatusWord := 4, [1,8].Status := 4, [1,8].OutputAddress := 43, [1,8].AlarmTimer.PRE := 2000, [1,8].AlarmTimerSP := 2, [1,8].AutoCloseTimer.ACC := 1104, [1,9].Tag := 'XV421', [1,9].CloseStatus := 1, [1,9].ZSOverride := 1, [1,9].EnableCfg := 1, [1,9].StatusWord := 4, [1,9].Status := 4,
        [1,9].OutputAddress := 44, [1,9].AlarmTimer.PRE := 2000, [1,9].AlarmTimerSP := 2, [1,9].AutoCloseTimer.ACC := 1105, [1,10].Tag := 'XV431', [1,10].CloseStatus := 1, [1,10].ZSOverride := 1, [1,10].EnableCfg := 1, [1,10].StatusWord := 4, [1,10].Status := 4, [1,10].OutputAddress := 45, [1,10].AlarmTimer.PRE := 2000, [1,10].AlarmTimerSP := 2, [1,10].AutoCloseTimer.ACC := 1104, [1,11].Tag := 'XV441', [1,11].CloseStatus := 1, [1,11].ZSOverride := 1, [1,11].EnableCfg := 1, [1,11].StatusWord := 4, [1,11].Status := 4, [1,11].OutputAddress := 46, [1,11].AlarmTimer.PRE := 2000, [1,11].AlarmTimerSP := 2, [1,11].AutoCloseTimer.ACC := 1103, [1,12].Tag := 'XV501', [1,12].CloseStatus := 1, [1,12].ZSOverride := 1, [1,12].EnableCfg := 1, [1,12].StatusWord := 4, [1,12].Status := 4, [1,12].OutputAddress := 39, [1,12].AlarmTimer.PRE := 2000, [1,12].AlarmTimerSP := 2, [1,12].AutoCloseTimer.ACC := 1072, [1,13].Tag := 'XV502', [1,13].CloseStatus := 1, [1,13].ZSOverride := 1, [1,13].EnableCfg := 1, [1,13].StatusWord := 4, [1,13].Status := 4, [1,13].OutputAddress := 40, [1,13].AlarmTimer.PRE := 2000, [1,13].AlarmTimerSP := 2, [1,13].AutoCloseTimer.ACC := 1016, [1,14].Tag := 'XV901', [1,14].CloseStatus := 1, [1,14].ZSOverride := 1, [1,14].EnableCfg := 1, [1,14].StatusWord := 4, [1,14].Status := 4, [1,14].OutputAddress := 37, [1,14].AlarmTimer.PRE := 2000, [1,14].AlarmTimerSP := 2, [1,15].OpenStatus := 1, [1,15].ZSOverride := 1, [1,15].OutputAddress := 47, [1,15].AlarmTimer.PRE := 2000, [1,15].AlarmTimerSP := 2, [1,16].CloseStatus := 1, [1,16].ZSOverride := 1,
        [1,16].OutputAddress := 48, [1,16].AlarmTimer.PRE := 2000, [1,16].AlarmTimerSP := 2, [1,17].OpenStatus := 1, [1,17].ZSOverride := 1, [1,17].OutputAddress := 49, [1,17].AlarmTimer.PRE := 2000, [1,17].AlarmTimerSP := 2, [1,17].AutoCloseTimer.ACC := 1594, [1,18].CloseStatus := 1, [1,18].ZSOverride := 1, [1,18].OutputAddress := 50, [1,18].AlarmTimer.PRE := 2000, [1,18].AlarmTimerSP := 2, [1,18].AutoCloseTimer.ACC := 137, [1,19].CloseStatus := 1, [1,19].ZSOverride := 1, [1,19].FailState := 1, [1,19].OutputAddress := 51, [1,19].AlarmTimer.PRE := 2000, [1,19].AlarmTimerSP := 2, [1,19].AutoCloseTimer.ACC := 1007, [1,20].CloseStatus := 1, [1,20].ZSOverride := 1, [1,20].OutputAddress := 52, [1,20].AlarmTimer.PRE := 2000, [1,20].AlarmTimerSP := 2, [1,20].AutoCloseTimer.ACC := 1004, [1,21].OpenStatus := 1, [1,21].ZSOverride := 1, [1,21].FailState := 1, [1,21].OutputAddress := 53, [1,21].AlarmTimer.PRE := 2000, [1,21].AlarmTimerSP := 2, [1,22].CloseStatus := 1, [1,22].ZSOverride := 1, [1,22].OutputAddress := 54, [1,22].AlarmTimer.PRE := 2000, [1,22].AlarmTimerSP := 2, [1,22].AutoCloseTimer.ACC := 131, [1,23].CloseStatus := 1, [1,23].ZSOverride := 1, [1,23].OutputAddress := 55, [1,23].AlarmTimer.PRE := 2000, [1,23].AlarmTimerSP := 2, [1,23].AutoCloseTimer.ACC := 1003, [1,24].CloseStatus := 1, [1,24].ZSOverride := 1, [1,24].OutputAddress := 56, [1,24].AlarmTimer.PRE := 2000, [1,24].AlarmTimerSP := 2, [1,24].AutoCloseTimer.ACC := 1002, [1,25].CloseStatus := 1, [1,25].ZSOverride := 1, [1,25].OutputAddress := 57, [1,25].AlarmTimer.PRE := 2000, [1,25].AlarmTimerSP := 2, [1,25].AutoCloseTimer.ACC := 1002, [1,26].CloseStatus := 1, [1,26].ZSOverride := 1,
        [1,26].OutputAddress := 58, [1,26].AlarmTimer.PRE := 2000, [1,26].AlarmTimerSP := 2, [1,26].AutoCloseTimer.ACC := 1002, [1,27].CloseStatus := 1, [1,27].ZSOverride := 1, [1,27].OutputAddress := 59, [1,27].AlarmTimer.PRE := 2000, [1,27].AlarmTimerSP := 2, [1,28].CloseStatus := 1, [1,28].ZSOverride := 1, [1,28].OutputAddress := 60, [1,28].AlarmTimer.PRE := 2000, [1,28].AlarmTimerSP := 2, [1,29].OpenStatus := 1, [1,29].ZSOverride := 1, [1,29].FailState := 1, [1,29].OutputAddress := 61, [1,29].AlarmTimer.PRE := 2000, [1,29].AlarmTimerSP := 2, [1,29].AutoCloseTimer.ACC := 1068, [1,30].CloseStatus := 1, [1,30].ZSOverride := 1, [1,30].OutputAddress := 62, [1,30].AlarmTimer.PRE := 2000, [1,30].AlarmTimerSP := 2, [1,30].AutoCloseTimer.ACC := 1069, [1,31].CloseStatus := 1, [1,31].ZSOverride := 1, [1,31].OutputAddress := 63, [1,31].AlarmTimer.PRE := 2000, [1,31].AlarmTimerSP := 2, [1,31].AutoCloseTimer.ACC := 131, [1,32].CloseStatus := 1, [1,32].PriorityCfg := 1, [1,32].ZSOpenAddress := 32, [1,32].OutputAddress := 68, [1,32].AlarmTimer.PRE := 2000, [1,32].AlarmTimerSP := 2, [1,32].AutoCloseTimer.ACC := 1059, [1,33].OpenStatus := 1, [1,33].PriorityCfg := 1, [1,33].FailState := 1, [1,33].ZSCloseAddress := 33, [1,33].OutputAddress := 69, [1,33].AlarmTimer.PRE := 2000, [1,33].AlarmTimerSP := 2, [1,33].AutoCloseTimer.ACC := 1123, [1,34].OpenStatus := 1, [1,34].PriorityCfg := 1, [1,34].FailState := 1, [1,34].ZSCloseAddress := 34, [1,34].OutputAddress := 70, [1,34].AlarmTimer.PRE := 2000, [1,34].AlarmTimerSP := 2, [1,34].AutoCloseTimer.ACC := 1095, [1,35].OpenStatus := 1, [1,35].PriorityCfg := 1, [1,35].FailState := 1, [1,35].ZSCloseAddress := 35,
        [1,35].OutputAddress := 71, [1,35].AlarmTimer.PRE := 2000, [1,35].AlarmTimerSP := 2, [1,35].AutoCloseTimer.ACC := 1127, [1,36].OpenStatus := 1, [1,36].PriorityCfg := 1, [1,36].FailState := 1, [1,36].ZSCloseAddress := 36, [1,36].OutputAddress := 72, [1,36].AlarmTimer.PRE := 2000, [1,36].AlarmTimerSP := 2, [1,36].AutoCloseTimer.ACC := 1004, [1,37].CloseStatus := 1, [1,37].PriorityCfg := 1, [1,37].ZSOpenAddress := 37, [1,37].OutputAddress := 73, [1,37].AlarmTimer.PRE := 2000, [1,37].AlarmTimerSP := 2, [1,37].AutoCloseTimer.ACC := 1121, [1,38].CloseStatus := 1, [1,38].Priority := 1, [1,38].PriorityCfg := 1, [1,38].ZSOpenAddress := 38, [1,38].OutputAddress := 40, [1,38].AlarmTimer.PRE := 2000, [1,38].AlarmTimerSP := 2, [1,38].AutoCloseTimer.ACC := 1135, [1,39].CloseStatus := 1, [1,39].Priority := 1, [1,39].PriorityCfg := 1, [1,39].ZSOpenAddress := 39, [1,39].OutputAddress := 41, [1,39].AlarmTimer.PRE := 2000, [1,39].AlarmTimerSP := 2, [1,39].AutoCloseTimer.ACC := 1121, [1,40].CloseStatus := 1, [1,40].Priority := 1, [1,40].PriorityCfg := 1, [1,40].ZSOpenAddress := 40, [1,40].OutputAddress := 42, [1,40].AlarmTimer.PRE := 2000, [1,40].AlarmTimerSP := 2, [1,40].AutoCloseTimer.ACC := 1112, [1,41].CloseStatus := 1, [1,41].Priority := 1, [1,41].PriorityCfg := 1, [1,41].ZSOpenAddress := 41, [1,41].OutputAddress := 43, [1,41].AlarmTimer.PRE := 2000, [1,41].AlarmTimerSP := 2, [1,42].CloseStatus := 1, [1,42].Priority := 1, [1,42].PriorityCfg := 1, [1,42].ZSOpenAddress := 42, [1,42].OutputAddress := 44, [1,42].AlarmTimer.PRE := 2000, [1,42].AlarmTimerSP := 2, [1,43].CloseStatus := 1, [1,43].Priority := 1, [1,43].PriorityCfg := 1,
        [1,43].ZSOpenAddress := 43, [1,43].OutputAddress := 52, [1,43].AlarmTimer.PRE := 2000, [1,43].AlarmTimerSP := 2, [1,44].CloseStatus := 1, [1,44].Priority := 1, [1,44].PriorityCfg := 1, [1,44].ZSOpenAddress := 44, [1,44].OutputAddress := 53, [1,44].AlarmTimer.PRE := 2000, [1,44].AlarmTimerSP := 2, [1,45].CloseStatus := 1, [1,45].Priority := 1, [1,45].PriorityCfg := 1, [1,45].ZSOpenAddress := 45, [1,45].OutputAddress := 54, [1,45].AlarmTimer.PRE := 2000, [1,45].AlarmTimerSP := 2, [1,46].CloseStatus := 1, [1,46].Priority := 1, [1,46].PriorityCfg := 1, [1,46].ZSOpenAddress := 46, [1,46].OutputAddress := 55, [1,46].AlarmTimer.PRE := 2000, [1,46].AlarmTimerSP := 2, [1,47].OpenStatus := 1, [1,47].Priority := 1, [1,47].PriorityCfg := 1, [1,47].FailState := 1, [1,47].ZSCloseAddress := 47, [1,47].OutputAddress := 45, [1,47].AlarmTimer.PRE := 2000, [1,47].AlarmTimerSP := 2, [1,48].FailState := 1, [1,48].ZSCloseAddress := 48, [1,48].OutputAddress := 80, [1,49].FailState := 1, [1,49].ZSCloseAddress := 49, [1,49].OutputAddress := 81, [1,50].FailState := 1, [1,50].ZSCloseAddress := 50, [1,50].OutputAddress := 82, [1,51].OpenStatus := 1, [1,51].FailState := 1, [1,51].ZSCloseAddress := 51, [1,51].OutputAddress := 83, [1,52].OpenStatus := 1, [1,52].FailState := 1, [1,52].ZSCloseAddress := 52, [1,52].OutputAddress := 84, [1,53].CloseStatus := 1, [1,53].FailState := 1, [1,53].ZSCloseAddress := 53, [1,53].OutputAddress := 85, [1,54].CloseStatus := 1, [1,54].FailState := 1, [1,54].ZSCloseAddress := 54, [1,54].OutputAddress := 86, [1,55].CloseStatus := 1, [1,55].FailState := 1,
        [1,55].ZSCloseAddress := 55, [1,55].OutputAddress := 87, [1,56].CloseStatus := 1, [1,58].CloseStatus := 1, [1,59].CloseStatus := 1, [2,0].Tag := 'XV001', [2,0].Control := 1, [2,0].Auto := 1, [2,0].Manual := 1, [2,0].OpenStatus := 1, [2,0].ZSOverride := 1, [2,0].FailState := 1, [2,0].EnableCfg := 1, [2,0].StatusWord := 2, [2,0].Status := 2, [2,0].OutputAddress := 32, [2,0].AlarmTimer.PRE := 2000, [2,0].AlarmTimerSP := 2, [2,1].Tag := 'XV002', [2,1].Control := 1, [2,1].Auto := 1, [2,1].Manual := 1, [2,1].OpenStatus := 1, [2,1].ZSOverride := 1, [2,1].FailState := 1, [2,1].EnableCfg := 1, [2,1].StatusWord := 2, [2,1].Status := 2, [2,1].OutputAddress := 33, [2,1].AlarmTimer.PRE := 2000, [2,1].AlarmTimerSP := 2, [2,1].AutoCloseTimer.ACC := 1103, [2,2].Tag := 'XV003', [2,2].CloseStatus := 1, [2,2].ZSOverride := 1, [2,2].EnableCfg := 1, [2,2].StatusWord := 4, [2,2].Status := 4, [2,2].OutputAddress := 34, [2,2].AlarmTimer.PRE := 2000, [2,2].AlarmTimerSP := 2, [2,2].AutoCloseTimer.ACC := 1032, [2,3].Tag := 'XV004', [2,3].Control := 1, [2,3].Auto := 1, [2,3].Manual := 1, [2,3].OpenStatus := 1, [2,3].ZSOverride := 1, [2,3].FailState := 1, [2,3].EnableCfg := 1, [2,3].StatusWord := 2, [2,3].Status := 2, [2,3].OutputAddress := 35, [2,3].AlarmTimer.PRE := 2000, [2,3].AlarmTimerSP := 2, [2,3].AutoCloseTimer.ACC := 1115, [2,4].Tag := 'XV005', [2,4].CloseStatus := 1, [2,4].ZSOverride := 1, [2,4].EnableCfg := 1,
        [2,4].StatusWord := 4, [2,4].Status := 4, [2,4].OutputAddress := 36, [2,4].AlarmTimer.PRE := 2000, [2,4].AlarmTimerSP := 2, [2,4].AutoCloseTimer.ACC := 1104, [2,5].Tag := 'XV102', [2,5].CloseStatus := 1, [2,5].ZSOverride := 1, [2,5].EnableCfg := 1, [2,5].StatusWord := 4, [2,5].Status := 4, [2,5].OutputAddress := 38, [2,5].AlarmTimer.PRE := 2000, [2,5].AlarmTimerSP := 2, [2,5].AutoCloseTimer.ACC := 1104, [2,6].Tag := 'XV401', [2,6].CloseStatus := 1, [2,6].ZSOverride := 1, [2,6].EnableCfg := 1, [2,6].StatusWord := 4, [2,6].Status := 4, [2,6].OutputAddress := 41, [2,6].AlarmTimer.PRE := 2000, [2,6].AlarmTimerSP := 2, [2,6].AutoCloseTimer.ACC := 1104, [2,7].Tag := 'XV402', [2,7].CloseStatus := 1, [2,7].ZSOverride := 1, [2,7].EnableCfg := 1, [2,7].StatusWord := 4, [2,7].Status := 4, [2,7].OutputAddress := 42, [2,7].AlarmTimer.PRE := 2000, [2,7].AlarmTimerSP := 2, [2,7].AutoCloseTimer.ACC := 1104, [2,8].Tag := 'XV411', [2,8].CloseStatus := 1, [2,8].EnableCfg := 1, [2,8].StatusWord := 4, [2,8].Status := 4, [2,8].OutputAddress := 43, [2,8].AlarmTimer.PRE := 2000, [2,8].AlarmTimerSP := 2, [2,8].AutoCloseTimer.ACC := 1104, [2,9].Tag := 'XV421', [2,9].CloseStatus := 1, [2,9].ZSOverride := 1, [2,9].EnableCfg := 1, [2,9].StatusWord := 4, [2,9].Status := 4, [2,9].OutputAddress := 44, [2,9].AlarmTimer.PRE := 2000, [2,9].AlarmTimerSP := 2, [2,9].AutoCloseTimer.ACC := 1105, [2,10].Tag := 'XV431', [2,10].CloseStatus := 1, [2,10].ZSOverride := 1, [2,10].EnableCfg := 1, [2,10].StatusWord := 4,
        [2,10].Status := 4, [2,10].OutputAddress := 45, [2,10].AlarmTimer.PRE := 2000, [2,10].AlarmTimerSP := 2, [2,10].AutoCloseTimer.ACC := 1104, [2,11].Tag := 'XV441', [2,11].CloseStatus := 1, [2,11].ZSOverride := 1, [2,11].EnableCfg := 1, [2,11].StatusWord := 4, [2,11].Status := 4, [2,11].OutputAddress := 46, [2,11].AlarmTimer.PRE := 2000, [2,11].AlarmTimerSP := 2, [2,11].AutoCloseTimer.ACC := 1103, [2,12].Tag := 'XV501', [2,12].CloseStatus := 1, [2,12].ZSOverride := 1, [2,12].StatusWord := 4, [2,12].Status := 4, [2,12].OutputAddress := 39, [2,12].AlarmTimer.PRE := 2000, [2,12].AlarmTimerSP := 2, [2,12].AutoCloseTimer.ACC := 1072, [2,13].Tag := 'XV502', [2,13].CloseStatus := 1, [2,13].ZSOverride := 1, [2,13].StatusWord := 4, [2,13].Status := 4, [2,13].OutputAddress := 40, [2,13].AlarmTimer.PRE := 2000, [2,13].AlarmTimerSP := 2, [2,13].AutoCloseTimer.ACC := 1016, [2,14].Tag := 'XV901', [2,14].CloseStatus := 1, [2,14].ZSOverride := 1, [2,14].EnableCfg := 1, [2,14].StatusWord := 4, [2,14].Status := 4, [2,14].OutputAddress := 37, [2,14].AlarmTimer.PRE := 2000, [2,14].AlarmTimerSP := 2, [2,15].OpenStatus := 1, [2,15].ZSOverride := 1, [2,15].FailState := 1, [2,15].OutputAddress := 47, [2,15].AlarmTimer.PRE := 2000, [2,15].AlarmTimerSP := 2, [2,16].CloseStatus := 1, [2,16].ZSOverride := 1, [2,16].OutputAddress := 48, [2,16].AlarmTimer.PRE := 2000, [2,16].AlarmTimerSP := 2, [2,17].OpenStatus := 1, [2,17].ZSOverride := 1, [2,17].FailState := 1, [2,17].OutputAddress := 49, [2,17].AlarmTimer.PRE := 2000, [2,17].AlarmTimerSP := 2, [2,17].AutoCloseTimer.ACC := 1594,
        [2,18].CloseStatus := 1, [2,18].ZSOverride := 1, [2,18].OutputAddress := 50, [2,18].AlarmTimer.PRE := 2000, [2,18].AlarmTimerSP := 2, [2,18].AutoCloseTimer.ACC := 137, [2,19].CloseStatus := 1, [2,19].ZSOverride := 1, [2,19].OutputAddress := 51, [2,19].AlarmTimer.PRE := 2000, [2,19].AlarmTimerSP := 2, [2,19].AutoCloseTimer.ACC := 1007, [2,20].CloseStatus := 1, [2,20].ZSOverride := 1, [2,20].OutputAddress := 52, [2,20].AlarmTimer.PRE := 2000, [2,20].AlarmTimerSP := 2, [2,20].AutoCloseTimer.ACC := 1004, [2,21].OpenStatus := 1, [2,21].ZSOverride := 1, [2,21].FailState := 1, [2,21].OutputAddress := 53, [2,21].AlarmTimer.PRE := 2000, [2,21].AlarmTimerSP := 2, [2,22].CloseStatus := 1, [2,22].ZSOverride := 1, [2,22].OutputAddress := 54, [2,22].AlarmTimer.PRE := 2000, [2,22].AlarmTimerSP := 2, [2,22].AutoCloseTimer.ACC := 131, [2,23].CloseStatus := 1, [2,23].ZSOverride := 1, [2,23].OutputAddress := 55, [2,23].AlarmTimer.PRE := 2000, [2,23].AlarmTimerSP := 2, [2,23].AutoCloseTimer.ACC := 1003, [2,24].CloseStatus := 1, [2,24].ZSOverride := 1, [2,24].OutputAddress := 56, [2,24].AlarmTimer.PRE := 2000, [2,24].AlarmTimerSP := 2, [2,24].AutoCloseTimer.ACC := 1002, [2,25].CloseStatus := 1, [2,25].ZSOverride := 1, [2,25].OutputAddress := 57, [2,25].AlarmTimer.PRE := 2000, [2,25].AlarmTimerSP := 2, [2,25].AutoCloseTimer.ACC := 1002, [2,26].CloseStatus := 1, [2,26].ZSOverride := 1, [2,26].OutputAddress := 58, [2,26].AlarmTimer.PRE := 2000, [2,26].AlarmTimerSP := 2, [2,26].AutoCloseTimer.ACC := 1002, [2,27].CloseStatus := 1, [2,27].ZSOverride := 1, [2,27].OutputAddress := 59, [2,27].AlarmTimer.PRE := 2000, [2,27].AlarmTimerSP := 2, [2,28].CloseStatus := 1,
        [2,28].ZSOverride := 1, [2,28].OutputAddress := 60, [2,28].AlarmTimer.PRE := 2000, [2,28].AlarmTimerSP := 2, [2,29].OpenStatus := 1, [2,29].ZSOverride := 1, [2,29].FailState := 1, [2,29].OutputAddress := 61, [2,29].AlarmTimer.PRE := 2000, [2,29].AlarmTimerSP := 2, [2,29].AutoCloseTimer.ACC := 1068, [2,30].CloseStatus := 1, [2,30].ZSOverride := 1, [2,30].OutputAddress := 62, [2,30].AlarmTimer.PRE := 2000, [2,30].AlarmTimerSP := 2, [2,30].AutoCloseTimer.ACC := 1069, [2,31].CloseStatus := 1, [2,31].ZSOverride := 1, [2,31].OutputAddress := 63, [2,31].AlarmTimer.PRE := 2000, [2,31].AlarmTimerSP := 2, [2,31].AutoCloseTimer.ACC := 131, [2,32].CloseStatus := 1, [2,32].PriorityCfg := 1, [2,32].AlarmTimerSP := 2, [2,32].AutoCloseTimer.ACC := 1059, [2,33].OpenStatus := 1, [2,33].PriorityCfg := 1, [2,33].AlarmTimerSP := 2, [2,33].AutoCloseTimer.ACC := 1123, [2,34].OpenStatus := 1, [2,34].PriorityCfg := 1, [2,34].AlarmTimerSP := 2, [2,34].AutoCloseTimer.ACC := 1095, [2,35].OpenStatus := 1, [2,35].PriorityCfg := 1, [2,35].AlarmTimerSP := 2, [2,35].AutoCloseTimer.ACC := 1127, [2,36].OpenStatus := 1, [2,36].PriorityCfg := 1, [2,36].AlarmTimerSP := 2, [2,36].AutoCloseTimer.ACC := 1004, [2,37].CloseStatus := 1, [2,37].PriorityCfg := 1, [2,37].AlarmTimerSP := 2, [2,37].AutoCloseTimer.ACC := 1121, [2,38].CloseStatus := 1, [2,38].Priority := 1, [2,38].PriorityCfg := 1, [2,38].AlarmTimerSP := 2, [2,38].AutoCloseTimer.ACC := 1135, [2,39].CloseStatus := 1, [2,39].Priority := 1, [2,39].PriorityCfg := 1, [2,39].AlarmTimerSP := 2, [2,39].AutoCloseTimer.ACC := 1121, [2,40].CloseStatus := 1, [2,40].Priority := 1, [2,40].PriorityCfg := 1,
        [2,40].AlarmTimerSP := 2, [2,40].AutoCloseTimer.ACC := 1112, [2,41].CloseStatus := 1, [2,41].Priority := 1, [2,41].PriorityCfg := 1, [2,41].AlarmTimerSP := 2, [2,42].CloseStatus := 1, [2,42].Priority := 1, [2,42].PriorityCfg := 1, [2,42].AlarmTimerSP := 2, [2,43].CloseStatus := 1, [2,43].Priority := 1, [2,43].PriorityCfg := 1, [2,43].AlarmTimerSP := 2, [2,44].CloseStatus := 1, [2,44].Priority := 1, [2,44].PriorityCfg := 1, [2,44].AlarmTimerSP := 2, [2,45].CloseStatus := 1, [2,45].Priority := 1, [2,45].PriorityCfg := 1, [2,45].AlarmTimerSP := 2, [2,46].CloseStatus := 1, [2,46].Priority := 1, [2,46].PriorityCfg := 1, [2,46].AlarmTimerSP := 2, [2,47].OpenStatus := 1, [2,47].Priority := 1, [2,47].PriorityCfg := 1, [2,47].AlarmTimerSP := 2, [2,51].OpenStatus := 1, [2,52].OpenStatus := 1, [2,53].CloseStatus := 1, [2,54].CloseStatus := 1, [2,55].CloseStatus := 1, [2,56].CloseStatus := 1, [2,58].CloseStatus := 1, [2,59].CloseStatus := 1, [3,0].CloseStatus := 1, [3,0].EnableCfg := 1, [3,0].StatusWord := 4, [3,0].Status := 4, [3,0].OutputAddress := 32, [3,1].CloseStatus := 1, [3,1].EnableCfg := 1, [3,1].StatusWord := 4, [3,1].Status := 4, [3,1].OutputAddress := 33, [3,2].CloseStatus := 1, [3,2].EnableCfg := 1, [3,2].StatusWord := 4, [3,2].Status := 4, [3,2].OutputAddress := 34, [3,3].CloseStatus := 1, [3,3].EnableCfg := 1, [3,3].StatusWord := 4, [3,3].Status := 4, [3,3].OutputAddress := 35, [3,4].CloseStatus := 1, [3,4].EnableCfg := 1,
        [3,4].StatusWord := 4, [3,4].Status := 4, [3,4].OutputAddress := 36, [3,5].CloseStatus := 1, [3,5].EnableCfg := 1, [3,5].StatusWord := 4, [3,5].Status := 4, [3,5].OutputAddress := 37, [3,6].CloseStatus := 1, [3,6].EnableCfg := 1, [3,6].StatusWord := 4, [3,6].Status := 4, [3,6].OutputAddress := 38, [3,7].CloseStatus := 1, [3,7].EnableCfg := 1, [3,7].StatusWord := 4, [3,7].Status := 4, [3,7].OutputAddress := 39, [3,8].CloseStatus := 1, [3,8].EnableCfg := 1, [3,8].StatusWord := 4, [3,8].Status := 4, [3,8].OutputAddress := 40, [3,9].CloseStatus := 1, [3,9].EnableCfg := 1, [3,9].StatusWord := 4, [3,9].Status := 4, [3,9].OutputAddress := 41, [3,10].CloseStatus := 1, [3,10].EnableCfg := 1, [3,10].StatusWord := 4, [3,10].Status := 4, [3,10].OutputAddress := 42, [3,11].CloseStatus := 1, [3,11].FailState := 1, [3,11].EnableCfg := 1, [3,11].StatusWord := 4, [3,11].Status := 4, [3,11].OutputAddress := 43, [3,12].CloseStatus := 1, [3,12].FailState := 1, [3,12].EnableCfg := 1, [3,12].StatusWord := 4, [3,12].Status := 4, [3,12].OutputAddress := 44, [3,13].CloseStatus := 1, [3,13].FailState := 1, [3,13].EnableCfg := 1, [3,13].StatusWord := 4, [3,13].Status := 4, [3,13].OutputAddress := 45, [3,14].CloseStatus := 1, [3,14].EnableCfg := 1, [3,14].StatusWord := 4, [3,14].Status := 4, [3,14].OutputAddress := 46, [3,15].CloseStatus := 1, [3,15].FailState := 1, [3,15].EnableCfg := 1, [3,15].StatusWord := 4,
        [3,15].Status := 4, [3,15].OutputAddress := 47, [3,16].CloseStatus := 1, [3,16].EnableCfg := 1, [3,16].StatusWord := 4, [3,16].Status := 4, [3,16].OutputAddress := 48, [3,17].CloseStatus := 1, [3,17].FailState := 1, [3,17].EnableCfg := 1, [3,17].StatusWord := 4, [3,17].Status := 4, [3,17].OutputAddress := 49, [3,18].CloseStatus := 1, [3,18].EnableCfg := 1, [3,18].StatusWord := 4, [3,18].Status := 4, [3,18].OutputAddress := 50, [3,19].CloseStatus := 1, [3,19].EnableCfg := 1, [3,19].StatusWord := 4, [3,19].Status := 4, [3,19].OutputAddress := 51, [3,20].CloseStatus := 1, [3,20].EnableCfg := 1, [3,20].StatusWord := 4, [3,20].Status := 4, [3,20].OutputAddress := 52, [3,21].CloseStatus := 1, [3,21].FailState := 1, [3,21].EnableCfg := 1, [3,21].StatusWord := 4, [3,21].Status := 4, [3,21].OutputAddress := 53, [3,22].CloseStatus := 1, [3,22].EnableCfg := 1, [3,22].StatusWord := 4, [3,22].Status := 4, [3,22].OutputAddress := 54, [3,23].CloseStatus := 1, [3,23].EnableCfg := 1, [3,23].StatusWord := 4, [3,23].Status := 4, [3,23].OutputAddress := 55, [3,24].CloseStatus := 1, [3,24].EnableCfg := 1, [3,24].StatusWord := 4, [3,24].Status := 4, [3,24].OutputAddress := 56, [3,25].CloseStatus := 1, [3,25].EnableCfg := 1, [3,25].StatusWord := 4, [3,25].Status := 4, [3,25].OutputAddress := 57, [3,26].CloseStatus := 1, [3,26].EnableCfg := 1, [3,26].StatusWord := 4, [3,26].Status := 4, [3,26].OutputAddress := 58, [3,27].CloseStatus := 1,
        [3,27].EnableCfg := 1, [3,27].StatusWord := 4, [3,27].Status := 4, [3,27].OutputAddress := 59, [3,28].CloseStatus := 1, [3,28].EnableCfg := 1, [3,28].StatusWord := 4, [3,28].Status := 4, [3,28].OutputAddress := 60, [3,29].CloseStatus := 1, [3,29].FailState := 1, [3,29].EnableCfg := 1, [3,29].StatusWord := 4, [3,29].Status := 4, [3,29].OutputAddress := 61, [3,30].CloseStatus := 1, [3,30].EnableCfg := 1, [3,30].StatusWord := 4, [3,30].Status := 4, [3,30].OutputAddress := 62, [3,31].CloseStatus := 1, [3,31].EnableCfg := 1, [3,31].StatusWord := 4, [3,31].Status := 4, [3,31].OutputAddress := 63, [4,0].Tag := 'XV001', [4,0].CloseStatus := 1, [4,0].ZSOverride := 1, [4,0].EnableCfg := 1, [4,0].StatusWord := 4, [4,0].Status := 4, [4,0].OutputAddress := 32, [4,0].AlarmTimer.PRE := 2000, [4,0].AlarmTimerSP := 2, [4,1].Tag := 'XV002', [4,1].CloseStatus := 1, [4,1].ZSOverride := 1, [4,1].EnableCfg := 1, [4,1].StatusWord := 4, [4,1].Status := 4, [4,1].OutputAddress := 33, [4,1].AlarmTimer.PRE := 2000, [4,1].AlarmTimerSP := 2, [4,1].AutoCloseTimer.ACC := 1103, [4,2].Tag := 'XV003', [4,2].CloseStatus := 1, [4,2].ZSOverride := 1, [4,2].EnableCfg := 1, [4,2].StatusWord := 4, [4,2].Status := 4, [4,2].OutputAddress := 34, [4,2].AlarmTimer.PRE := 2000, [4,2].AlarmTimerSP := 2, [4,2].AutoCloseTimer.ACC := 1032, [4,3].Tag := 'XV004', [4,3].CloseStatus := 1, [4,3].ZSOverride := 1, [4,3].EnableCfg := 1, [4,3].StatusWord := 4, [4,3].Status := 4,
        [4,3].OutputAddress := 35, [4,3].AlarmTimer.PRE := 2000, [4,3].AlarmTimerSP := 2, [4,3].AutoCloseTimer.ACC := 1115, [4,4].Tag := 'XV005', [4,4].CloseStatus := 1, [4,4].ZSOverride := 1, [4,4].EnableCfg := 1, [4,4].StatusWord := 4, [4,4].Status := 4, [4,4].OutputAddress := 36, [4,4].AlarmTimer.PRE := 2000, [4,4].AlarmTimerSP := 2, [4,4].AutoCloseTimer.ACC := 1104, [4,5].Tag := 'XV006', [4,5].CloseStatus := 1, [4,5].ZSOverride := 1, [4,5].EnableCfg := 1, [4,5].StatusWord := 4, [4,5].Status := 4, [4,5].OutputAddress := 37, [4,5].AlarmTimer.PRE := 2000, [4,5].AlarmTimerSP := 2, [4,5].AutoCloseTimer.ACC := 1104, [4,6].Tag := 'XV007', [4,6].CloseStatus := 1, [4,6].ZSOverride := 1, [4,6].EnableCfg := 1, [4,6].StatusWord := 4, [4,6].Status := 4, [4,6].OutputAddress := 38, [4,6].AlarmTimer.PRE := 2000, [4,6].AlarmTimerSP := 2, [4,6].AutoCloseTimer.ACC := 1104, [4,7].Tag := 'XV008', [4,7].CloseStatus := 1, [4,7].ZSOverride := 1, [4,7].EnableCfg := 1, [4,7].StatusWord := 4, [4,7].Status := 4, [4,7].OutputAddress := 39, [4,7].AlarmTimer.PRE := 2000, [4,7].AlarmTimerSP := 2, [4,7].AutoCloseTimer.ACC := 1104, [4,8].Tag := 'XV009', [4,8].CloseStatus := 1, [4,8].ZSOverride := 1, [4,8].EnableCfg := 1, [4,8].StatusWord := 4, [4,8].Status := 4, [4,8].OutputAddress := 40, [4,8].AlarmTimer.PRE := 2000, [4,8].AlarmTimerSP := 2, [4,8].AutoCloseTimer.ACC := 1104, [4,9].Tag := 'XV010', [4,9].CloseStatus := 1, [4,9].ZSOverride := 1, [4,9].EnableCfg := 1, [4,9].StatusWord := 4, [4,9].Status := 4,
        [4,9].OutputAddress := 41, [4,9].AlarmTimer.PRE := 2000, [4,9].AlarmTimerSP := 2, [4,9].AutoCloseTimer.ACC := 1105, [4,10].Tag := 'XV011', [4,10].CloseStatus := 1, [4,10].ZSOverride := 1, [4,10].EnableCfg := 1, [4,10].StatusWord := 4, [4,10].Status := 4, [4,10].OutputAddress := 42, [4,10].AlarmTimer.PRE := 2000, [4,10].AlarmTimerSP := 2, [4,10].AutoCloseTimer.ACC := 1104, [4,11].Tag := 'XV012', [4,11].Control := 1, [4,11].Auto := 1, [4,11].Manual := 1, [4,11].OpenStatus := 1, [4,11].ZSOverride := 1, [4,11].FailState := 1, [4,11].EnableCfg := 1, [4,11].StatusWord := 2, [4,11].Status := 2, [4,11].OutputAddress := 43, [4,11].AlarmTimer.PRE := 2000, [4,11].AlarmTimerSP := 2, [4,11].AutoCloseTimer.ACC := 1103, [4,12].Tag := 'XV013', [4,12].Control := 1, [4,12].Auto := 1, [4,12].Manual := 1, [4,12].OpenStatus := 1, [4,12].ZSOverride := 1, [4,12].FailState := 1, [4,12].EnableCfg := 1, [4,12].StatusWord := 2, [4,12].Status := 2, [4,12].OutputAddress := 44, [4,12].AlarmTimer.PRE := 2000, [4,12].AlarmTimerSP := 2, [4,12].AutoCloseTimer.ACC := 1072, [4,13].Tag := 'XV014', [4,13].Control := 1, [4,13].Auto := 1, [4,13].Manual := 1, [4,13].OpenStatus := 1, [4,13].ZSOverride := 1, [4,13].FailState := 1, [4,13].EnableCfg := 1, [4,13].StatusWord := 2, [4,13].Status := 2, [4,13].OutputAddress := 45, [4,13].AlarmTimer.PRE := 2000, [4,13].AlarmTimerSP := 2, [4,13].AutoCloseTimer.ACC := 1016, [4,14].Tag := 'XV015', [4,14].CloseStatus := 1, [4,14].ZSOverride := 1, [4,14].EnableCfg := 1,
        [4,14].StatusWord := 4, [4,14].Status := 4, [4,14].OutputAddress := 46, [4,14].AlarmTimer.PRE := 2000, [4,14].AlarmTimerSP := 2, [4,15].Tag := 'XV016', [4,15].Control := 1, [4,15].Auto := 1, [4,15].Manual := 1, [4,15].OpenStatus := 1, [4,15].ZSOverride := 1, [4,15].FailState := 1, [4,15].EnableCfg := 1, [4,15].StatusWord := 2, [4,15].Status := 2, [4,15].OutputAddress := 47, [4,15].AlarmTimer.PRE := 2000, [4,15].AlarmTimerSP := 2, [4,16].Tag := 'XV017', [4,16].CloseStatus := 1, [4,16].ZSOverride := 1, [4,16].EnableCfg := 1, [4,16].StatusWord := 4, [4,16].Status := 4, [4,16].OutputAddress := 48, [4,16].AlarmTimer.PRE := 2000, [4,16].AlarmTimerSP := 2, [4,17].Tag := 'XV018', [4,17].Control := 1, [4,17].Auto := 1, [4,17].Manual := 1, [4,17].OpenStatus := 1, [4,17].ZSOverride := 1, [4,17].FailState := 1, [4,17].EnableCfg := 1, [4,17].StatusWord := 2, [4,17].Status := 2, [4,17].OutputAddress := 49, [4,17].AlarmTimer.PRE := 2000, [4,17].AlarmTimerSP := 2, [4,17].AutoCloseTimer.ACC := 1594, [4,18].Tag := 'XV019', [4,18].CloseStatus := 1, [4,18].ZSOverride := 1, [4,18].EnableCfg := 1, [4,18].StatusWord := 4, [4,18].Status := 4, [4,18].OutputAddress := 50, [4,18].AlarmTimer.PRE := 2000, [4,18].AlarmTimerSP := 2, [4,18].AutoCloseTimer.ACC := 137, [4,19].Tag := 'XV020', [4,19].CloseStatus := 1, [4,19].ZSOverride := 1, [4,19].EnableCfg := 1, [4,19].StatusWord := 4, [4,19].Status := 4, [4,19].OutputAddress := 51, [4,19].AlarmTimer.PRE := 2000, [4,19].AlarmTimerSP := 2,
        [4,19].AutoCloseTimer.ACC := 1007, [4,20].Tag := 'XV021', [4,20].CloseStatus := 1, [4,20].ZSOverride := 1, [4,20].EnableCfg := 1, [4,20].StatusWord := 4, [4,20].Status := 4, [4,20].OutputAddress := 52, [4,20].AlarmTimer.PRE := 2000, [4,20].AlarmTimerSP := 2, [4,20].AutoCloseTimer.ACC := 1004, [4,21].Tag := 'XV022', [4,21].Control := 1, [4,21].Auto := 1, [4,21].Manual := 1, [4,21].OpenStatus := 1, [4,21].ZSOverride := 1, [4,21].FailState := 1, [4,21].EnableCfg := 1, [4,21].StatusWord := 2, [4,21].Status := 2, [4,21].OutputAddress := 53, [4,21].AlarmTimer.PRE := 2000, [4,21].AlarmTimerSP := 2, [4,22].Tag := 'XV023', [4,22].CloseStatus := 1, [4,22].ZSOverride := 1, [4,22].EnableCfg := 1, [4,22].StatusWord := 4, [4,22].Status := 4, [4,22].OutputAddress := 54, [4,22].AlarmTimer.PRE := 2000, [4,22].AlarmTimerSP := 2, [4,22].AutoCloseTimer.ACC := 131, [4,23].Tag := 'XV024', [4,23].CloseStatus := 1, [4,23].ZSOverride := 1, [4,23].EnableCfg := 1, [4,23].StatusWord := 4, [4,23].Status := 4, [4,23].OutputAddress := 55, [4,23].AlarmTimer.PRE := 2000, [4,23].AlarmTimerSP := 2, [4,23].AutoCloseTimer.ACC := 1003, [4,24].Tag := 'XV025', [4,24].CloseStatus := 1, [4,24].ZSOverride := 1, [4,24].EnableCfg := 1, [4,24].StatusWord := 4, [4,24].Status := 4, [4,24].OutputAddress := 56, [4,24].AlarmTimer.PRE := 2000, [4,24].AlarmTimerSP := 2, [4,24].AutoCloseTimer.ACC := 1002, [4,25].Tag := 'XV026', [4,25].CloseStatus := 1, [4,25].ZSOverride := 1, [4,25].EnableCfg := 1, [4,25].StatusWord := 4, [4,25].Status := 4,
        [4,25].OutputAddress := 57, [4,25].AlarmTimer.PRE := 2000, [4,25].AlarmTimerSP := 2, [4,25].AutoCloseTimer.ACC := 1002, [4,26].Tag := 'XV028', [4,26].CloseStatus := 1, [4,26].ZSOverride := 1, [4,26].EnableCfg := 1, [4,26].StatusWord := 4, [4,26].Status := 4, [4,26].OutputAddress := 58, [4,26].AlarmTimer.PRE := 2000, [4,26].AlarmTimerSP := 2, [4,26].AutoCloseTimer.ACC := 1002, [4,27].Tag := 'XV029', [4,27].CloseStatus := 1, [4,27].ZSOverride := 1, [4,27].EnableCfg := 1, [4,27].StatusWord := 4, [4,27].Status := 4, [4,27].OutputAddress := 59, [4,27].AlarmTimer.PRE := 2000, [4,27].AlarmTimerSP := 2, [4,28].Tag := 'XV030', [4,28].CloseStatus := 1, [4,28].ZSOverride := 1, [4,28].EnableCfg := 1, [4,28].StatusWord := 4, [4,28].Status := 4, [4,28].OutputAddress := 60, [4,28].AlarmTimer.PRE := 2000, [4,28].AlarmTimerSP := 2, [4,29].Tag := 'XV031', [4,29].Control := 1, [4,29].Auto := 1, [4,29].Manual := 1, [4,29].OpenStatus := 1, [4,29].ZSOverride := 1, [4,29].FailState := 1, [4,29].EnableCfg := 1, [4,29].StatusWord := 2, [4,29].Status := 2, [4,29].OutputAddress := 61, [4,29].AlarmTimer.PRE := 2000, [4,29].AlarmTimerSP := 2, [4,29].AutoCloseTimer.ACC := 1068, [4,30].Tag := 'XV033', [4,30].CloseStatus := 1, [4,30].ZSOverride := 1, [4,30].EnableCfg := 1, [4,30].StatusWord := 4, [4,30].Status := 4, [4,30].OutputAddress := 62, [4,30].AlarmTimer.PRE := 2000, [4,30].AlarmTimerSP := 2, [4,30].AutoCloseTimer.ACC := 1069, [4,31].Tag := 'XV034', [4,31].CloseStatus := 1, [4,31].ZSOverride := 1, [4,31].EnableCfg := 1,
        [4,31].StatusWord := 4, [4,31].Status := 4, [4,31].OutputAddress := 63, [4,31].AlarmTimer.PRE := 2000, [4,31].AlarmTimerSP := 2, [4,31].AutoCloseTimer.ACC := 131, [4,32].CloseStatus := 1, [4,32].PriorityCfg := 1, [4,32].ZSOpenAddress := 32, [4,32].OutputAddress := 68, [4,32].AlarmTimer.PRE := 2000, [4,32].AlarmTimerSP := 2, [4,32].AutoCloseTimer.ACC := 1059, [4,33].OpenStatus := 1, [4,33].PriorityCfg := 1, [4,33].FailState := 1, [4,33].ZSCloseAddress := 33, [4,33].OutputAddress := 69, [4,33].AlarmTimer.PRE := 2000, [4,33].AlarmTimerSP := 2, [4,33].AutoCloseTimer.ACC := 1123, [4,34].OpenStatus := 1, [4,34].PriorityCfg := 1, [4,34].FailState := 1, [4,34].ZSCloseAddress := 34, [4,34].OutputAddress := 70, [4,34].AlarmTimer.PRE := 2000, [4,34].AlarmTimerSP := 2, [4,34].AutoCloseTimer.ACC := 1095, [4,35].OpenStatus := 1, [4,35].PriorityCfg := 1, [4,35].FailState := 1, [4,35].ZSCloseAddress := 35, [4,35].OutputAddress := 71, [4,35].AlarmTimer.PRE := 2000, [4,35].AlarmTimerSP := 2, [4,35].AutoCloseTimer.ACC := 1127, [4,36].OpenStatus := 1, [4,36].PriorityCfg := 1, [4,36].FailState := 1, [4,36].ZSCloseAddress := 36, [4,36].OutputAddress := 72, [4,36].AlarmTimer.PRE := 2000, [4,36].AlarmTimerSP := 2, [4,36].AutoCloseTimer.ACC := 1004, [4,37].CloseStatus := 1, [4,37].PriorityCfg := 1, [4,37].ZSOpenAddress := 37, [4,37].OutputAddress := 73, [4,37].AlarmTimer.PRE := 2000, [4,37].AlarmTimerSP := 2, [4,37].AutoCloseTimer.ACC := 1121, [4,38].CloseStatus := 1, [4,38].Priority := 1, [4,38].PriorityCfg := 1, [4,38].ZSOpenAddress := 38, [4,38].OutputAddress := 40, [4,38].AlarmTimer.PRE := 2000, [4,38].AlarmTimerSP := 2, [4,38].AutoCloseTimer.ACC := 1135,
        [4,39].CloseStatus := 1, [4,39].Priority := 1, [4,39].PriorityCfg := 1, [4,39].ZSOpenAddress := 39, [4,39].OutputAddress := 41, [4,39].AlarmTimer.PRE := 2000, [4,39].AlarmTimerSP := 2, [4,39].AutoCloseTimer.ACC := 1121, [4,40].CloseStatus := 1, [4,40].Priority := 1, [4,40].PriorityCfg := 1, [4,40].ZSOpenAddress := 40, [4,40].OutputAddress := 42, [4,40].AlarmTimer.PRE := 2000, [4,40].AlarmTimerSP := 2, [4,40].AutoCloseTimer.ACC := 1112, [4,41].CloseStatus := 1, [4,41].Priority := 1, [4,41].PriorityCfg := 1, [4,41].ZSOpenAddress := 41, [4,41].OutputAddress := 43, [4,41].AlarmTimer.PRE := 2000, [4,41].AlarmTimerSP := 2, [4,42].CloseStatus := 1, [4,42].Priority := 1, [4,42].PriorityCfg := 1, [4,42].ZSOpenAddress := 42, [4,42].OutputAddress := 44, [4,42].AlarmTimer.PRE := 2000, [4,42].AlarmTimerSP := 2, [4,43].CloseStatus := 1, [4,43].Priority := 1, [4,43].PriorityCfg := 1, [4,43].ZSOpenAddress := 43, [4,43].OutputAddress := 52, [4,43].AlarmTimer.PRE := 2000, [4,43].AlarmTimerSP := 2, [4,44].CloseStatus := 1, [4,44].Priority := 1, [4,44].PriorityCfg := 1, [4,44].ZSOpenAddress := 44, [4,44].OutputAddress := 53, [4,44].AlarmTimer.PRE := 2000, [4,44].AlarmTimerSP := 2, [4,45].CloseStatus := 1, [4,45].Priority := 1, [4,45].PriorityCfg := 1, [4,45].ZSOpenAddress := 45, [4,45].OutputAddress := 54, [4,45].AlarmTimer.PRE := 2000, [4,45].AlarmTimerSP := 2, [4,46].CloseStatus := 1, [4,46].Priority := 1, [4,46].PriorityCfg := 1, [4,46].ZSOpenAddress := 46, [4,46].OutputAddress := 55, [4,46].AlarmTimer.PRE := 2000, [4,46].AlarmTimerSP := 2, [4,47].OpenStatus := 1, [4,47].Priority := 1,
        [4,47].PriorityCfg := 1, [4,47].FailState := 1, [4,47].ZSCloseAddress := 47, [4,47].OutputAddress := 45, [4,47].AlarmTimer.PRE := 2000, [4,47].AlarmTimerSP := 2, [4,48].FailState := 1, [4,48].ZSCloseAddress := 48, [4,48].OutputAddress := 80, [4,49].FailState := 1, [4,49].ZSCloseAddress := 49, [4,49].OutputAddress := 81, [4,50].FailState := 1, [4,50].ZSCloseAddress := 50, [4,50].OutputAddress := 82, [4,51].OpenStatus := 1, [4,51].FailState := 1, [4,51].ZSCloseAddress := 51, [4,51].OutputAddress := 83, [4,52].OpenStatus := 1, [4,52].FailState := 1, [4,52].ZSCloseAddress := 52, [4,52].OutputAddress := 84, [4,53].CloseStatus := 1, [4,53].FailState := 1, [4,53].ZSCloseAddress := 53, [4,53].OutputAddress := 85, [4,54].CloseStatus := 1, [4,54].FailState := 1, [4,54].ZSCloseAddress := 54, [4,54].OutputAddress := 86, [4,55].CloseStatus := 1, [4,55].FailState := 1, [4,55].ZSCloseAddress := 55, [4,55].OutputAddress := 87, [4,56].CloseStatus := 1, [4,58].CloseStatus := 1, [4,59].CloseStatus := 1, [5,0].Tag := 'XV001', [5,0].CloseStatus := 1, [5,0].ZSOverride := 1, [5,0].EnableCfg := 1, [5,0].StatusWord := 4, [5,0].Status := 4, [5,0].OutputAddress := 32, [5,0].AlarmTimer.PRE := 2000, [5,0].AlarmTimerSP := 2, [5,1].Tag := 'XV002', [5,1].CloseStatus := 1, [5,1].ZSOverride := 1, [5,1].EnableCfg := 1, [5,1].StatusWord := 4, [5,1].Status := 4, [5,1].OutputAddress := 33, [5,1].AlarmTimer.PRE := 2000, [5,1].AlarmTimerSP := 2, [5,1].AutoCloseTimer.ACC := 1103, [5,2].Tag := 'XV003', [5,2].CloseStatus := 1, [5,2].ZSOverride := 1,
        [5,2].EnableCfg := 1, [5,2].StatusWord := 4, [5,2].Status := 4, [5,2].OutputAddress := 34, [5,2].AlarmTimer.PRE := 2000, [5,2].AlarmTimerSP := 2, [5,2].AutoCloseTimer.ACC := 1032, [5,3].Tag := 'XV004', [5,3].CloseStatus := 1, [5,3].ZSOverride := 1, [5,3].EnableCfg := 1, [5,3].StatusWord := 4, [5,3].Status := 4, [5,3].OutputAddress := 35, [5,3].AlarmTimer.PRE := 2000, [5,3].AlarmTimerSP := 2, [5,3].AutoCloseTimer.ACC := 1115, [5,4].Tag := 'XV005', [5,4].CloseStatus := 1, [5,4].ZSOverride := 1, [5,4].EnableCfg := 1, [5,4].StatusWord := 4, [5,4].Status := 4, [5,4].OutputAddress := 36, [5,4].AlarmTimer.PRE := 2000, [5,4].AlarmTimerSP := 2, [5,4].AutoCloseTimer.ACC := 1104, [5,5].Tag := 'XV006', [5,5].CloseStatus := 1, [5,5].ZSOverride := 1, [5,5].EnableCfg := 1, [5,5].StatusWord := 4, [5,5].Status := 4, [5,5].OutputAddress := 37, [5,5].AlarmTimer.PRE := 2000, [5,5].AlarmTimerSP := 2, [5,5].AutoCloseTimer.ACC := 1104, [5,6].Tag := 'XV007', [5,6].CloseStatus := 1, [5,6].ZSOverride := 1, [5,6].EnableCfg := 1, [5,6].StatusWord := 4, [5,6].Status := 4, [5,6].OutputAddress := 38, [5,6].AlarmTimer.PRE := 2000, [5,6].AlarmTimerSP := 2, [5,6].AutoCloseTimer.ACC := 1104, [5,7].Tag := 'XV008', [5,7].CloseStatus := 1, [5,7].ZSOverride := 1, [5,7].EnableCfg := 1, [5,7].StatusWord := 4, [5,7].Status := 4, [5,7].OutputAddress := 39, [5,7].AlarmTimer.PRE := 2000, [5,7].AlarmTimerSP := 2, [5,7].AutoCloseTimer.ACC := 1104, [5,8].Tag := 'XV009', [5,8].CloseStatus := 1, [5,8].ZSOverride := 1,
        [5,8].EnableCfg := 1, [5,8].StatusWord := 4, [5,8].Status := 4, [5,8].OutputAddress := 40, [5,8].AlarmTimer.PRE := 2000, [5,8].AlarmTimerSP := 2, [5,8].AutoCloseTimer.ACC := 1104, [5,9].Tag := 'XV010', [5,9].CloseStatus := 1, [5,9].ZSOverride := 1, [5,9].EnableCfg := 1, [5,9].StatusWord := 4, [5,9].Status := 4, [5,9].OutputAddress := 41, [5,9].AlarmTimer.PRE := 2000, [5,9].AlarmTimerSP := 2, [5,9].AutoCloseTimer.ACC := 1105, [5,10].Tag := 'XV011', [5,10].CloseStatus := 1, [5,10].ZSOverride := 1, [5,10].EnableCfg := 1, [5,10].StatusWord := 4, [5,10].Status := 4, [5,10].OutputAddress := 42, [5,10].AlarmTimer.PRE := 2000, [5,10].AlarmTimerSP := 2, [5,10].AutoCloseTimer.ACC := 1104, [5,11].Tag := 'XV012', [5,11].Control := 1, [5,11].Auto := 1, [5,11].Manual := 1, [5,11].OpenStatus := 1, [5,11].ZSOverride := 1, [5,11].FailState := 1, [5,11].EnableCfg := 1, [5,11].StatusWord := 2, [5,11].Status := 2, [5,11].OutputAddress := 43, [5,11].AlarmTimer.PRE := 2000, [5,11].AlarmTimerSP := 2, [5,11].AutoCloseTimer.ACC := 1103, [5,12].Tag := 'XV013', [5,12].Control := 1, [5,12].Auto := 1, [5,12].Manual := 1, [5,12].OpenStatus := 1, [5,12].ZSOverride := 1, [5,12].FailState := 1, [5,12].EnableCfg := 1, [5,12].StatusWord := 2, [5,12].Status := 2, [5,12].OutputAddress := 44, [5,12].AlarmTimer.PRE := 2000, [5,12].AlarmTimerSP := 2, [5,12].AutoCloseTimer.ACC := 1072, [5,13].Tag := 'XV014', [5,13].Control := 1, [5,13].Auto := 1, [5,13].Manual := 1, [5,13].OpenStatus := 1,
        [5,13].ZSOverride := 1, [5,13].FailState := 1, [5,13].EnableCfg := 1, [5,13].StatusWord := 2, [5,13].Status := 2, [5,13].OutputAddress := 45, [5,13].AlarmTimer.PRE := 2000, [5,13].AlarmTimerSP := 2, [5,13].AutoCloseTimer.ACC := 1016, [5,14].Tag := 'XV015', [5,14].CloseStatus := 1, [5,14].ZSOverride := 1, [5,14].EnableCfg := 1, [5,14].StatusWord := 4, [5,14].Status := 4, [5,14].OutputAddress := 46, [5,14].AlarmTimer.PRE := 2000, [5,14].AlarmTimerSP := 2, [5,15].Tag := 'XV016', [5,15].Control := 1, [5,15].Auto := 1, [5,15].Manual := 1, [5,15].OpenStatus := 1, [5,15].ZSOverride := 1, [5,15].FailState := 1, [5,15].EnableCfg := 1, [5,15].StatusWord := 2, [5,15].Status := 2, [5,15].OutputAddress := 47, [5,15].AlarmTimer.PRE := 2000, [5,15].AlarmTimerSP := 2, [5,16].Tag := 'XV017', [5,16].CloseStatus := 1, [5,16].ZSOverride := 1, [5,16].EnableCfg := 1, [5,16].StatusWord := 4, [5,16].Status := 4, [5,16].OutputAddress := 48, [5,16].AlarmTimer.PRE := 2000, [5,16].AlarmTimerSP := 2, [5,17].Tag := 'XV018', [5,17].Control := 1, [5,17].Auto := 1, [5,17].Manual := 1, [5,17].OpenStatus := 1, [5,17].ZSOverride := 1, [5,17].FailState := 1, [5,17].EnableCfg := 1, [5,17].StatusWord := 2, [5,17].Status := 2, [5,17].OutputAddress := 49, [5,17].AlarmTimer.PRE := 2000, [5,17].AlarmTimerSP := 2, [5,17].AutoCloseTimer.ACC := 1594, [5,18].Tag := 'XV019', [5,18].CloseStatus := 1, [5,18].ZSOverride := 1, [5,18].EnableCfg := 1, [5,18].StatusWord := 4, [5,18].Status := 4,
        [5,18].OutputAddress := 50, [5,18].AlarmTimer.PRE := 2000, [5,18].AlarmTimerSP := 2, [5,18].AutoCloseTimer.ACC := 137, [5,19].Tag := 'XV020', [5,19].CloseStatus := 1, [5,19].ZSOverride := 1, [5,19].EnableCfg := 1, [5,19].StatusWord := 4, [5,19].Status := 4, [5,19].OutputAddress := 51, [5,19].AlarmTimer.PRE := 2000, [5,19].AlarmTimerSP := 2, [5,19].AutoCloseTimer.ACC := 1007, [5,20].Tag := 'XV021', [5,20].CloseStatus := 1, [5,20].ZSOverride := 1, [5,20].EnableCfg := 1, [5,20].StatusWord := 4, [5,20].Status := 4, [5,20].OutputAddress := 52, [5,20].AlarmTimer.PRE := 2000, [5,20].AlarmTimerSP := 2, [5,20].AutoCloseTimer.ACC := 1004, [5,21].Tag := 'XV022', [5,21].Control := 1, [5,21].Auto := 1, [5,21].Manual := 1, [5,21].OpenStatus := 1, [5,21].ZSOverride := 1, [5,21].FailState := 1, [5,21].EnableCfg := 1, [5,21].StatusWord := 2, [5,21].Status := 2, [5,21].OutputAddress := 53, [5,21].AlarmTimer.PRE := 2000, [5,21].AlarmTimerSP := 2, [5,22].Tag := 'XV023', [5,22].CloseStatus := 1, [5,22].ZSOverride := 1, [5,22].EnableCfg := 1, [5,22].StatusWord := 4, [5,22].Status := 4, [5,22].OutputAddress := 54, [5,22].AlarmTimer.PRE := 2000, [5,22].AlarmTimerSP := 2, [5,22].AutoCloseTimer.ACC := 131, [5,23].Tag := 'XV024', [5,23].CloseStatus := 1, [5,23].ZSOverride := 1, [5,23].EnableCfg := 1, [5,23].StatusWord := 4, [5,23].Status := 4, [5,23].OutputAddress := 55, [5,23].AlarmTimer.PRE := 2000, [5,23].AlarmTimerSP := 2, [5,23].AutoCloseTimer.ACC := 1003, [5,24].Tag := 'XV025', [5,24].CloseStatus := 1, [5,24].ZSOverride := 1,
        [5,24].EnableCfg := 1, [5,24].StatusWord := 4, [5,24].Status := 4, [5,24].OutputAddress := 56, [5,24].AlarmTimer.PRE := 2000, [5,24].AlarmTimerSP := 2, [5,24].AutoCloseTimer.ACC := 1002, [5,25].Tag := 'XV026', [5,25].CloseStatus := 1, [5,25].ZSOverride := 1, [5,25].EnableCfg := 1, [5,25].StatusWord := 4, [5,25].Status := 4, [5,25].OutputAddress := 57, [5,25].AlarmTimer.PRE := 2000, [5,25].AlarmTimerSP := 2, [5,25].AutoCloseTimer.ACC := 1002, [5,26].Tag := 'XV028', [5,26].CloseStatus := 1, [5,26].ZSOverride := 1, [5,26].EnableCfg := 1, [5,26].StatusWord := 4, [5,26].Status := 4, [5,26].OutputAddress := 58, [5,26].AlarmTimer.PRE := 2000, [5,26].AlarmTimerSP := 2, [5,26].AutoCloseTimer.ACC := 1002, [5,27].Tag := 'XV029', [5,27].CloseStatus := 1, [5,27].ZSOverride := 1, [5,27].EnableCfg := 1, [5,27].StatusWord := 4, [5,27].Status := 4, [5,27].OutputAddress := 59, [5,27].AlarmTimer.PRE := 2000, [5,27].AlarmTimerSP := 2, [5,28].Tag := 'XV030', [5,28].CloseStatus := 1, [5,28].ZSOverride := 1, [5,28].EnableCfg := 1, [5,28].StatusWord := 4, [5,28].Status := 4, [5,28].OutputAddress := 60, [5,28].AlarmTimer.PRE := 2000, [5,28].AlarmTimerSP := 2, [5,29].Tag := 'XV031', [5,29].Control := 1, [5,29].Auto := 1, [5,29].Manual := 1, [5,29].OpenStatus := 1, [5,29].ZSOverride := 1, [5,29].FailState := 1, [5,29].EnableCfg := 1, [5,29].StatusWord := 2, [5,29].Status := 2, [5,29].OutputAddress := 61, [5,29].AlarmTimer.PRE := 2000, [5,29].AlarmTimerSP := 2, [5,29].AutoCloseTimer.ACC := 1068, [5,30].Tag := 'XV033',
        [5,30].CloseStatus := 1, [5,30].ZSOverride := 1, [5,30].EnableCfg := 1, [5,30].StatusWord := 4, [5,30].Status := 4, [5,30].OutputAddress := 62, [5,30].AlarmTimer.PRE := 2000, [5,30].AlarmTimerSP := 2, [5,30].AutoCloseTimer.ACC := 1069, [5,31].Tag := 'XV034', [5,31].CloseStatus := 1, [5,31].ZSOverride := 1, [5,31].EnableCfg := 1, [5,31].StatusWord := 4, [5,31].Status := 4, [5,31].OutputAddress := 63, [5,31].AlarmTimer.PRE := 2000, [5,31].AlarmTimerSP := 2, [5,31].AutoCloseTimer.ACC := 131, [5,32].CloseStatus := 1, [5,32].PriorityCfg := 1, [5,32].ZSOpenAddress := 32, [5,32].OutputAddress := 68, [5,32].AlarmTimer.PRE := 2000, [5,32].AlarmTimerSP := 2, [5,32].AutoCloseTimer.ACC := 1059, [5,33].OpenStatus := 1, [5,33].PriorityCfg := 1, [5,33].FailState := 1, [5,33].ZSCloseAddress := 33, [5,33].OutputAddress := 69, [5,33].AlarmTimer.PRE := 2000, [5,33].AlarmTimerSP := 2, [5,33].AutoCloseTimer.ACC := 1123, [5,34].OpenStatus := 1, [5,34].PriorityCfg := 1, [5,34].FailState := 1, [5,34].ZSCloseAddress := 34, [5,34].OutputAddress := 70, [5,34].AlarmTimer.PRE := 2000, [5,34].AlarmTimerSP := 2, [5,34].AutoCloseTimer.ACC := 1095, [5,35].OpenStatus := 1, [5,35].PriorityCfg := 1, [5,35].FailState := 1, [5,35].ZSCloseAddress := 35, [5,35].OutputAddress := 71, [5,35].AlarmTimer.PRE := 2000, [5,35].AlarmTimerSP := 2, [5,35].AutoCloseTimer.ACC := 1127, [5,36].OpenStatus := 1, [5,36].PriorityCfg := 1, [5,36].FailState := 1, [5,36].ZSCloseAddress := 36, [5,36].OutputAddress := 72, [5,36].AlarmTimer.PRE := 2000, [5,36].AlarmTimerSP := 2, [5,36].AutoCloseTimer.ACC := 1004, [5,37].CloseStatus := 1, [5,37].PriorityCfg := 1,
        [5,37].ZSOpenAddress := 37, [5,37].OutputAddress := 73, [5,37].AlarmTimer.PRE := 2000, [5,37].AlarmTimerSP := 2, [5,37].AutoCloseTimer.ACC := 1121, [5,38].CloseStatus := 1, [5,38].Priority := 1, [5,38].PriorityCfg := 1, [5,38].ZSOpenAddress := 38, [5,38].OutputAddress := 40, [5,38].AlarmTimer.PRE := 2000, [5,38].AlarmTimerSP := 2, [5,38].AutoCloseTimer.ACC := 1135, [5,39].CloseStatus := 1, [5,39].Priority := 1, [5,39].PriorityCfg := 1, [5,39].ZSOpenAddress := 39, [5,39].OutputAddress := 41, [5,39].AlarmTimer.PRE := 2000, [5,39].AlarmTimerSP := 2, [5,39].AutoCloseTimer.ACC := 1121, [5,40].CloseStatus := 1, [5,40].Priority := 1, [5,40].PriorityCfg := 1, [5,40].ZSOpenAddress := 40, [5,40].OutputAddress := 42, [5,40].AlarmTimer.PRE := 2000, [5,40].AlarmTimerSP := 2, [5,40].AutoCloseTimer.ACC := 1112, [5,41].CloseStatus := 1, [5,41].Priority := 1, [5,41].PriorityCfg := 1, [5,41].ZSOpenAddress := 41, [5,41].OutputAddress := 43, [5,41].AlarmTimer.PRE := 2000, [5,41].AlarmTimerSP := 2, [5,42].CloseStatus := 1, [5,42].Priority := 1, [5,42].PriorityCfg := 1, [5,42].ZSOpenAddress := 42, [5,42].OutputAddress := 44, [5,42].AlarmTimer.PRE := 2000, [5,42].AlarmTimerSP := 2, [5,43].CloseStatus := 1, [5,43].Priority := 1, [5,43].PriorityCfg := 1, [5,43].ZSOpenAddress := 43, [5,43].OutputAddress := 52, [5,43].AlarmTimer.PRE := 2000, [5,43].AlarmTimerSP := 2, [5,44].CloseStatus := 1, [5,44].Priority := 1, [5,44].PriorityCfg := 1, [5,44].ZSOpenAddress := 44, [5,44].OutputAddress := 53, [5,44].AlarmTimer.PRE := 2000, [5,44].AlarmTimerSP := 2, [5,45].CloseStatus := 1, [5,45].Priority := 1, [5,45].PriorityCfg := 1,
        [5,45].ZSOpenAddress := 45, [5,45].OutputAddress := 54, [5,45].AlarmTimer.PRE := 2000, [5,45].AlarmTimerSP := 2, [5,46].CloseStatus := 1, [5,46].Priority := 1, [5,46].PriorityCfg := 1, [5,46].ZSOpenAddress := 46, [5,46].OutputAddress := 55, [5,46].AlarmTimer.PRE := 2000, [5,46].AlarmTimerSP := 2, [5,47].OpenStatus := 1, [5,47].Priority := 1, [5,47].PriorityCfg := 1, [5,47].FailState := 1, [5,47].ZSCloseAddress := 47, [5,47].OutputAddress := 45, [5,47].AlarmTimer.PRE := 2000, [5,47].AlarmTimerSP := 2, [5,48].FailState := 1, [5,48].ZSCloseAddress := 48, [5,48].OutputAddress := 80, [5,49].FailState := 1, [5,49].ZSCloseAddress := 49, [5,49].OutputAddress := 81, [5,50].FailState := 1, [5,50].ZSCloseAddress := 50, [5,50].OutputAddress := 82, [5,51].OpenStatus := 1, [5,51].FailState := 1, [5,51].ZSCloseAddress := 51, [5,51].OutputAddress := 83, [5,52].OpenStatus := 1, [5,52].FailState := 1, [5,52].ZSCloseAddress := 52, [5,52].OutputAddress := 84, [5,53].CloseStatus := 1, [5,53].FailState := 1, [5,53].ZSCloseAddress := 53, [5,53].OutputAddress := 85, [5,54].CloseStatus := 1, [5,54].FailState := 1, [5,54].ZSCloseAddress := 54, [5,54].OutputAddress := 86, [5,55].CloseStatus := 1, [5,55].FailState := 1, [5,55].ZSCloseAddress := 55, [5,55].OutputAddress := 87, [5,56].CloseStatus := 1, [5,58].CloseStatus := 1, [5,59].CloseStatus := 1);
   ValveControl : ValveControl := (ValveStatus1 := 30847, MaxValveNum := 32);   // Valve Control
   ValveSwInput : BOOL[64];   // Valve digital input
   VersionLetterForDevelopment : STRING := '.b';   // Version Letter for Development
   VersionNumberForRelease : STRING := '3.02.00.00';   // Version Number for Release
   WI001 : ALIAS FOR AnalogPoint[15];   // Feed Bag Weight
   WI001_SIG : ALIAS FOR DigitalPoint[94];
   WI001Alarm : ALIAS FOR AlarmAnalog[15];   // Feed Bag Weight Alarm
   WI101 : ALIAS FOR AnalogPoint[0];   // Filtrate Weight
   WI101_SIG : ALIAS FOR DigitalPoint[95];
   WI101Alarm : ALIAS FOR AlarmAnalog[0];   // Filtrate Weight Alarm
   WI102 : ALIAS FOR AnalogPoint[1];   // Customer Filtrate Weight
   WI102_SIG : ALIAS FOR DigitalPoint[96];
   WI102Alarm : ALIAS FOR AlarmAnalog[1];   // Customer Filtrate Weight Alarm
   XC102_3 : ALIAS FOR DigitalOutput[5];   // UV Auto Zero
   XC102_3DF : ALIAS FOR DigitalPoint[13];   // C8000 Defect
   XS001 : ALIAS FOR DigitalPoint[1];   // Door Closed
   XS002 : ALIAS FOR DigitalPoint[6];   // Clamshell Locking 1 Closed
   XS003 : ALIAS FOR DigitalPoint[7];   // Clamshell Locking 2 Closed
   XS006 : ALIAS FOR DigitalPoint[2];   // Door to Frame Locking Closed
   XS011 : ALIAS FOR DigitalPoint[11];   // Pump P001 Type
   XS012 : ALIAS FOR DigitalPoint[12];   // Pump P002 Type
   XV001 : ALIAS FOR Valve[0];   // XV001
   XV002 : ALIAS FOR Valve[1];   // XV002
   XV003 : ALIAS FOR Valve[2];   // XV003
   XV004 : ALIAS FOR Valve[3];   // XV004
   XV005 : ALIAS FOR Valve[4];   // XV005
   XV006 : ALIAS FOR Valve[19];
   XV007 : ALIAS FOR Valve[20];
   XV102 : ALIAS FOR Valve[5];   // XV102
   XV401 : ALIAS FOR Valve[6];   // XV401
   XV402 : ALIAS FOR Valve[7];   // XV402
   XV403 : ALIAS FOR Valve[15];
   XV404 : ALIAS FOR Valve[16];
   XV405 : ALIAS FOR Valve[17];
   XV406 : ALIAS FOR Valve[18];
   XV411 : ALIAS FOR Valve[8];   // XV411
   XV421 : ALIAS FOR Valve[9];   // XV421
   XV431 : ALIAS FOR Valve[10];   // XV431
   XV441 : ALIAS FOR Valve[11];   // XV441
   XV501 : ALIAS FOR Valve[12];   // XV501
   XV502 : ALIAS FOR Valve[13];   // XV502
   XV901 : ALIAS FOR Valve[14];   // XV901
   Y500A : ALIAS FOR DigitalOutput[11];   // Unlock Clamshell
   Y500B : ALIAS FOR DigitalOutput[12];   // Lock Clamshell
   Y501A : ALIAS FOR DigitalOutput[10];   // Unlock Door
   Y501B : ALIAS FOR DigitalOutput[9];   // Lock Door
   Y502A : ALIAS FOR DigitalOutput[13];   // Unlock Clamshell in Door
   Y502B : ALIAS FOR DigitalOutput[14];   // Lock Clamshell in Door
   Y503A : ALIAS FOR DigitalOutput[15];   // Connect Clamshell
   Y503B : ALIAS FOR DigitalOutput[16];   // Disconnect Clamshell
   YA01 : ALIAS FOR DigitalPoint[50];   // PC to PLC communication failure
   YA02 : ALIAS FOR DigitalPoint[51];   // CCP Runtime communication failure
   YA03 : ALIAS FOR DigitalPoint[52];   // Historical Data collection failure
   YA04 : ALIAS FOR DigitalPoint[53];   // Hard Drive Overload
   YA05 : ALIAS FOR DigitalPoint[54];   // Database Overload
   YA06 : ALIAS FOR DigitalPoint[55];   // Node 0 communication failure - Smart
   YA07 : ALIAS FOR DigitalPoint[56];   // Node 0 internal defect - Smart
   YA08 : ALIAS FOR DigitalPoint[57];   // Node 1 communication failure - Clamshell
   YA09 : ALIAS FOR DigitalPoint[58];   // Node 1 internal defect - Clamshell
   YA10 : ALIAS FOR DigitalPoint[59];   // PLC Program Major Fault
   YA11 : ALIAS FOR DigitalPoint[60];   // Database Corrupted
   YA12 : ALIAS FOR DigitalPoint[61];   // Unauthorized accesses
   YA13 : ALIAS FOR DigitalPoint[62];   // Tank Size Mismatch
   YA14 : ALIAS FOR DigitalPoint[63];   // SQL Server Write Failure
   YA15 : ALIAS FOR DigitalPoint[69];   // Node 3 Communication Failure - Pump
   YA16 : ALIAS FOR DigitalPoint[70];   // Node 3 Internal Defect - Pump
   YA17 : ALIAS FOR DigitalPoint[71];   // Node 4 Communication Failure - Instrum
   YA18 : ALIAS FOR DigitalPoint[72];   // Node 4 Internal Defect - Instrum
   YA19 : ALIAS FOR DigitalPoint[73];   // Node 5 Communication Failure - Tank
   YA20 : ALIAS FOR DigitalPoint[74];   // Node 5 Internal Defect - Tank
   YA21 : ALIAS FOR DigitalPoint[75];   // Node 6 IND331 Communication Failure
   YA22 : ALIAS FOR DigitalPoint[76];   // Node 7 IND131 Communication Failure
   YA41 : ALIAS FOR DigitalPoint[77];   // YA41 Operating Time Exceeded
   ZSDF : ALIAS FOR DigitalPoint[68];   // ZSDF Clamshell Locking Defect
END_VAR
